--- program side_paint (robot ABB IRB 5500-27) ---
  Smooth(1)
  Set speed (1000.0 mm/s)
  Set Ref.: FrameSidePaint
  Set Tool: Paint gun
  Show Paint gun
  MoveJ 1 to (-1297.14, 952.77, 801.05) mm, rotated rx -98.58 ry 36.73 rz 174.5 deg; joints [-13.501, 53.284, -35.7, -53.192, 43.737, -41.413, -170]
  MoveL 2 to (-1297.14, 952.77, 801.05) mm, rotated rx -98.58 ry 36.73 rz 174.5 deg; joints [-13.501, 53.284, -35.7, -53.192, 43.737, -41.413, -170]
  MoveL 3 to (-1297.75, 853.49, 789.09) mm, rotated rx -98.58 ry 36.73 rz 174.5 deg; joints [-15.474, 56.036, -39.978, -51.479, 40.206, -40.518, -170]
  MoveL 4 to (-1297.75, 853.49, 789.09) mm, rotated rx -98.58 ry 36.73 rz 174.5 deg; joints [-15.474, 56.036, -39.978, -51.479, 40.206, -40.518, -170]
  Set speed (50.0 mm/s)
  MoveL 5 to (-1297.75, 853.39, 796.9) mm, rotated rx -98.58 ry 36.73 rz 174.5 deg; joints [-15.482, 55.905, -40.062, -50.968, 39.758, -40.731, -170]
  Set speed (1000.0 mm/s)
  MoveL 6 to (-1297.75, 853.39, 796.9) mm, rotated rx -98.58 ry 36.73 rz 174.5 deg; joints [-15.482, 55.905, -40.062, -50.968, 39.758, -40.731, -170]
  MoveL 7 to (-1297.14, 952.67, 808.86) mm, rotated rx -98.58 ry 36.73 rz 174.5 deg; joints [-13.509, 53.15, -35.783, -52.711, 43.305, -41.606, -170]
  Set speed (1000.0 mm/s)
  MoveL 8 to (-1377.47, 943.1, 874.94) mm, rotated rx -98.65 ry 38.29 rz 174.46 deg; joints [-14.496, 49.055, -31.026, -57.58, 47.073, -38.423, -170]
  MoveL 9 to (-1377.75, 843.8, 863.14) mm, rotated rx -98.65 ry 38.29 rz 174.46 deg; joints [-16.488, 51.747, -35.093, -56.497, 44.013, -37.161, -170]
  MoveL 10 to (-1377.75, 843.8, 863.14) mm, rotated rx -98.65 ry 38.29 rz 174.46 deg; joints [-16.488, 51.747, -35.093, -56.497, 44.013, -37.161, -170]
  Set speed (50.0 mm/s)
  MoveL 11 to (-1377.75, 845.82, 854.57) mm, rotated rx -98.73 ry 37.85 rz 174.4 deg; joints [-16.458, 51.746, -34.877, -56.091, 43.595, -37.432, -170]
  MoveL 12 to (-1377.75, 852.68, 825.37) mm, rotated rx -98.99 ry 36.5 rz 174.23 deg; joints [-16.347, 51.788, -34.184, -54.959, 42.475, -38.231, -170]
  MoveL 13 to (-1377.75, 852.68, 825.37) mm, rotated rx -98.99 ry 36.5 rz 174.23 deg; joints [-16.347, 51.788, -34.184, -54.959, 42.475, -38.231, -170]
  MoveL 14 to (-1377.75, 852.9, 804.32) mm, rotated rx -98.93 ry 36.57 rz 174.27 deg; joints [-16.325, 52.17, -33.954, -56.498, 43.866, -37.653, -170]
  MoveL 15 to (-1377.75, 853.2, 774.32) mm, rotated rx -98.85 ry 36.66 rz 174.33 deg; joints [-16.297, 52.733, -33.656, -58.588, 45.794, -36.9, -170]
  MoveL 16 to (-1377.75, 853.51, 744.32) mm, rotated rx -98.76 ry 36.76 rz 174.38 deg; joints [-16.27, 53.316, -33.393, -60.572, 47.664, -36.222, -170]
  MoveL 17 to (-1377.75, 853.62, 723.27) mm, rotated rx -96.67 ry 38.01 rz 175.72 deg; joints [-16.272, 54.302, -33.281, -66.947, 53.226, -34.784, -170]
  MoveL 18 to (-1377.75, 853.79, 693.27) mm, rotated rx -92.96 ry 22.32 rz 178.98 deg; joints [-17.183, 52.483, -31.27, -47.624, 27.861, -47.672, -170]
  MoveL 19 to (-1377.75, 853.95, 663.27) mm, rotated rx -90.24 ry 20.37 rz -179.71 deg; joints [-17.303, 53.259, -30.78, -52.353, 29.913, -47.74, -170]
  MoveL 20 to (-1377.75, 854, 636.95) mm, rotated rx -90.22 ry 20.39 rz -179.69 deg; joints [-17.278, 53.814, -30.63, -54.436, 31.655, -46.867, -170]
  MoveL 21 to (-1377.75, 854.06, 606.95) mm, rotated rx -90.19 ry 20.4 rz -179.67 deg; joints [-17.254, 54.461, -30.491, -56.636, 33.537, -45.983, -170]
  MoveL 22 to (-1377.75, 854.12, 576.95) mm, rotated rx -90.16 ry 20.41 rz -179.64 deg; joints [-17.232, 55.127, -30.383, -58.679, 35.325, -45.201, -170]
  MoveL 23 to (-1377.75, 854.18, 546.95) mm, rotated rx -90.13 ry 20.43 rz -179.62 deg; joints [-17.213, 55.809, -30.307, -60.585, 37.031, -44.505, -170]
  MoveL 24 to (-1377.75, 854.23, 516.95) mm, rotated rx -90.1 ry 20.44 rz -179.6 deg; joints [-17.195, 56.507, -30.263, -62.373, 38.664, -43.883, -170]
  MoveL 25 to (-1377.75, 854.25, 508.95) mm, rotated rx -90.1 ry 20.44 rz -179.6 deg; joints [-17.19, 56.695, -30.258, -62.801, 39.067, -43.739, -170]
  Set speed (1000.0 mm/s)
  MoveL 26 to (-1377.75, 854.25, 508.95) mm, rotated rx -90.1 ry 20.44 rz -179.6 deg; joints [-17.19, 56.695, -30.258, -62.801, 39.067, -43.739, -170]
  MoveL 27 to (-1378.51, 954.25, 509.11) mm, rotated rx -90.1 ry 20.44 rz -179.6 deg; joints [-15.183, 54.375, -26.133, -63.747, 42.417, -45.012, -170]
  Set speed (1000.0 mm/s)
  MoveL 28 to (-1458.68, 953.67, 187.25) mm, rotated rx -89.99 ry 0.54 rz -179.47 deg; joints [-16.728, 56.853, -21.556, -35.057, 15.198, -66.186, -170]
  MoveL 29 to (-1457.75, 853.67, 187.27) mm, rotated rx -89.99 ry 0.54 rz -179.47 deg; joints [-18.915, 58.968, -25.635, -25.442, 6.373, -70.654, -170]
  MoveL 30 to (-1457.75, 853.67, 187.27) mm, rotated rx -89.99 ry 0.54 rz -179.47 deg; joints [-18.915, 58.968, -25.635, -25.442, 6.373, -70.654, -170]
  Set speed (50.0 mm/s)
  MoveL 31 to (-1457.75, 853.67, 195.27) mm, rotated rx -89.99 ry 0.54 rz -179.47 deg; joints [-18.972, 58.745, -25.612, -22.234, 4.29, -72.531, -170]
  MoveL 32 to (-1457.75, 853.67, 225.27) mm, rotated rx -90 ry 20.52 rz -179.48 deg; joints [-18.06, 61.359, -26.112, -80.802, 56.365, -38.648, -170]
  MoveL 33 to (-1457.75, 853.67, 255.27) mm, rotated rx -90 ry 20.51 rz -179.49 deg; joints [-18.066, 60.5, -25.864, -79.807, 55.247, -38.783, -170]
  MoveL 34 to (-1457.75, 853.67, 285.27) mm, rotated rx -90.01 ry 20.51 rz -179.5 deg; joints [-18.073, 59.656, -25.644, -78.771, 54.095, -38.938, -170]
  MoveL 35 to (-1457.75, 853.67, 315.27) mm, rotated rx -90.01 ry 20.5 rz -179.51 deg; joints [-18.079, 58.826, -25.455, -77.693, 52.908, -39.114, -170]
  MoveL 36 to (-1457.75, 853.67, 345.27) mm, rotated rx -90.02 ry 20.49 rz -179.52 deg; joints [-18.087, 58.011, -25.294, -76.57, 51.684, -39.312, -170]
  MoveL 37 to (-1457.75, 853.67, 375.27) mm, rotated rx -90.02 ry 20.48 rz -179.53 deg; joints [-18.095, 57.21, -25.164, -75.399, 50.423, -39.536, -170]
  MoveL 38 to (-1457.75, 853.66, 405.27) mm, rotated rx -90.03 ry 20.48 rz -179.53 deg; joints [-18.104, 56.424, -25.062, -74.178, 49.125, -39.788, -170]
  MoveL 39 to (-1457.75, 853.66, 435.27) mm, rotated rx -90.03 ry 20.47 rz -179.54 deg; joints [-18.114, 55.652, -24.99, -72.903, 47.786, -40.071, -170]
  MoveL 40 to (-1457.75, 853.66, 465.27) mm, rotated rx -90.04 ry 20.46 rz -179.55 deg; joints [-18.124, 54.896, -24.946, -71.569, 46.405, -40.387, -170]
  MoveL 41 to (-1457.75, 853.66, 495.27) mm, rotated rx -90.04 ry 20.46 rz -179.56 deg; joints [-18.135, 54.155, -24.932, -70.172, 44.981, -40.741, -170]
  MoveL 42 to (-1457.75, 853.66, 526.08) mm, rotated rx -90.05 ry 20.45 rz -179.57 deg; joints [-18.148, 53.41, -24.949, -68.666, 43.469, -41.147, -170]
  MoveL 43 to (-1457.75, 853.62, 556.08) mm, rotated rx -90.07 ry 20.43 rz -179.59 deg; joints [-18.161, 52.696, -24.998, -67.057, 41.898, -41.604, -170]
  MoveL 44 to (-1457.75, 853.58, 586.08) mm, rotated rx -90.1 ry 20.42 rz -179.62 deg; joints [-18.176, 51.999, -25.077, -65.36, 40.27, -42.117, -170]
  MoveL 45 to (-1457.75, 853.52, 628.44) mm, rotated rx -90.14 ry 20.4 rz -179.65 deg; joints [-18.199, 51.042, -25.24, -62.791, 37.864, -42.951, -170]
  MoveL 46 to (-1457.75, 853.41, 658.44) mm, rotated rx -90.2 ry 20.38 rz -179.69 deg; joints [-18.219, 50.379, -25.397, -60.74, 36.008, -43.651, -170]
  MoveL 47 to (-1457.75, 853.3, 688.44) mm, rotated rx -90.25 ry 20.36 rz -179.73 deg; joints [-18.241, 49.734, -25.586, -58.544, 34.065, -44.447, -170]
  MoveL 48 to (-1457.75, 853.15, 730.8) mm, rotated rx -90.34 ry 20.33 rz -179.78 deg; joints [-18.277, 48.852, -25.907, -55.141, 31.145, -45.766, -170]
  MoveL 49 to (-1457.75, 852.89, 760.79) mm, rotated rx -92.62 ry 22.9 rz 179.1 deg; joints [-18.125, 48.27, -26.437, -53.114, 31.255, -44.471, -170]
  MoveL 50 to (-1457.75, 852.62, 790.79) mm, rotated rx -94.76 ry 18.59 rz 178.38 deg; joints [-18.675, 46.691, -27.128, -19.032, 6.195, -62.515, -170]
  MoveL 51 to (-1457.75, 852.24, 833.15) mm, rotated rx -99.29 ry 36.39 rz 174.04 deg; joints [-17.25, 48.344, -28.68, -59.788, 46.031, -35.543, -170]
  MoveL 52 to (-1457.75, 842.15, 874) mm, rotated rx -99.06 ry 37.76 rz 174.19 deg; joints [-17.436, 48.149, -29.605, -60.089, 46.37, -34.987, -170]
  MoveL 53 to (-1457.75, 832.57, 914.98) mm, rotated rx -98.75 ry 39.5 rz 174.39 deg; joints [-17.596, 48.056, -30.593, -61.046, 47.459, -34.165, -170]
  MoveL 54 to (-1457.75, 829.64, 928.8) mm, rotated rx -100.09 ry 40.17 rz 173.53 deg; joints [-17.613, 47.828, -31.021, -59.139, 46.443, -34.036, -170]
  Set speed (1000.0 mm/s)
  MoveL 55 to (-1457.75, 829.64, 928.8) mm, rotated rx -100.09 ry 40.17 rz 173.53 deg; joints [-17.613, 47.828, -31.021, -59.139, 46.443, -34.036, -170]
  MoveL 56 to (-1457.88, 928.74, 942.19) mm, rotated rx -100.09 ry 40.17 rz 173.53 deg; joints [-15.61, 45.122, -27.108, -59.778, 49.118, -35.52, -170]
  Set speed (1000.0 mm/s)
  MoveL 57 to (-1538.66, 913.21, 1014.54) mm, rotated rx -105.61 ry 41.62 rz 170.03 deg; joints [-16.814, 40.69, -24.051, -54.13, 45.376, -33.626, -170]
  MoveL 58 to (-1537.75, 815.25, 994.43) mm, rotated rx -105.61 ry 41.62 rz 170.03 deg; joints [-18.805, 43.502, -27.729, -53.938, 43.177, -32.043, -170]
  MoveL 59 to (-1537.75, 815.25, 994.43) mm, rotated rx -105.61 ry 41.62 rz 170.03 deg; joints [-18.805, 43.502, -27.729, -53.938, 43.177, -32.043, -170]
  Set speed (50.0 mm/s)
  MoveL 60 to (-1537.75, 817.42, 984.35) mm, rotated rx -105.7 ry 41.25 rz 169.97 deg; joints [-18.767, 43.525, -27.488, -53.735, 42.978, -32.204, -170]
  MoveL 61 to (-1537.75, 823.74, 955.02) mm, rotated rx -106.39 ry 38.88 rz 169.55 deg; joints [-18.708, 43.372, -26.899, -49.424, 39.023, -34.352, -170]
  MoveL 62 to (-1537.75, 830.36, 927.04) mm, rotated rx -102.94 ry 38.8 rz 171.73 deg; joints [-18.566, 44.073, -25.879, -57.39, 44.7, -32.92, -170]
  MoveL 63 to (-1537.75, 837.26, 897.85) mm, rotated rx -99.3 ry 38.2 rz 174.04 deg; joints [-18.489, 44.817, -24.916, -64.229, 49.447, -32.46, -170]
  MoveL 64 to (-1537.75, 844.38, 869.99) mm, rotated rx -99.44 ry 37.24 rz 173.95 deg; joints [-18.359, 44.951, -24.277, -64.056, 49.208, -32.848, -170]
  MoveL 65 to (-1537.75, 851.81, 840.93) mm, rotated rx -108.52 ry 36.78 rz 168.22 deg; joints [-18.104, 43.97, -24.492, -49.321, 40.009, -34.298, -170]
  MoveL 66 to (-1537.75, 852.15, 797.55) mm, rotated rx -101.05 ry 38.75 rz 172.92 deg; joints [-18.073, 46.114, -23.379, -67.854, 54.496, -30.798, -170]
  MoveL 67 to (-1537.75, 852.4, 767.56) mm, rotated rx -94.65 ry 21.55 rz 178.41 deg; joints [-19.181, 44.634, -21.632, -51.982, 29.331, -43.354, -170]
  MoveL 68 to (-1537.75, 852.64, 737.56) mm, rotated rx -90.09 ry 20.34 rz -179.69 deg; joints [-19.27, 45.923, -20.99, -62.422, 36.243, -42.294, -170]
  MoveL 69 to (-1537.75, 852.77, 694.18) mm, rotated rx -90.06 ry 20.37 rz -179.66 deg; joints [-19.242, 46.844, -20.673, -65.334, 38.948, -41.323, -170]
  MoveL 70 to (-1537.75, 852.86, 664.18) mm, rotated rx -90.04 ry 20.38 rz -179.63 deg; joints [-19.226, 47.501, -20.49, -67.203, 40.732, -40.746, -170]
  MoveL 71 to (-1537.75, 852.95, 634.18) mm, rotated rx -90.02 ry 20.4 rz -179.6 deg; joints [-19.211, 48.176, -20.337, -68.97, 42.453, -40.235, -170]
  MoveL 72 to (-1537.75, 852.98, 590.81) mm, rotated rx -90 ry 20.42 rz -179.58 deg; joints [-19.193, 49.178, -20.172, -71.312, 44.799, -39.612, -170]
  MoveL 73 to (-1537.75, 853.01, 560.81) mm, rotated rx -89.99 ry 20.44 rz -179.56 deg; joints [-19.181, 49.891, -20.094, -72.839, 46.362, -39.24, -170]
  MoveL 74 to (-1537.75, 853.03, 530.81) mm, rotated rx -89.98 ry 20.45 rz -179.55 deg; joints [-19.171, 50.619, -20.044, -74.297, 47.879, -38.91, -170]
  MoveL 75 to (-1537.75, 853.02, 496.12) mm, rotated rx -89.98 ry 20.46 rz -179.54 deg; joints [-19.16, 51.478, -20.025, -75.864, 49.547, -38.588, -170]
  MoveL 76 to (-1537.75, 853.02, 466.12) mm, rotated rx -89.98 ry 20.47 rz -179.53 deg; joints [-19.151, 52.238, -20.038, -77.16, 50.948, -38.345, -170]
  MoveL 77 to (-1537.75, 853.01, 436.12) mm, rotated rx -89.97 ry 20.47 rz -179.52 deg; joints [-19.143, 53.012, -20.08, -78.405, 52.311, -38.132, -170]
  MoveL 78 to (-1537.75, 853, 406.12) mm, rotated rx -89.97 ry 20.48 rz -179.51 deg; joints [-19.136, 53.8, -20.15, -79.602, 53.639, -37.945, -170]
  MoveL 79 to (-1537.75, 852.99, 376.12) mm, rotated rx -89.97 ry 20.49 rz -179.51 deg; joints [-19.129, 54.603, -20.249, -80.755, 54.932, -37.784, -170]
  MoveL 80 to (-1537.75, 852.98, 346.12) mm, rotated rx -89.97 ry 20.49 rz -179.5 deg; joints [-19.123, 55.42, -20.375, -81.866, 56.191, -37.645, -170]
  MoveL 81 to (-1537.75, 852.97, 316.12) mm, rotated rx -89.97 ry 20.5 rz -179.49 deg; joints [-19.117, 56.251, -20.529, -82.938, 57.418, -37.526, -170]
  MoveL 82 to (-1537.75, 852.96, 286.12) mm, rotated rx -89.97 ry 0.51 rz -179.49 deg; joints [-19.911, 53.732, -20.278, -31.164, 8.952, -66.908, -170]
  MoveL 83 to (-1537.75, 852.95, 256.12) mm, rotated rx -89.97 ry 0.52 rz -179.49 deg; joints [-19.811, 54.549, -20.328, -37.182, 13.072, -63.574, -170]
  MoveL 84 to (-1537.75, 852.94, 226.12) mm, rotated rx -89.97 ry 0.52 rz -179.48 deg; joints [-19.743, 55.38, -20.423, -41.507, 16.152, -61.281, -170]
  MoveL 85 to (-1537.75, 852.94, 196.12) mm, rotated rx -89.97 ry 0.53 rz -179.47 deg; joints [-19.691, 56.224, -20.555, -44.993, 18.721, -59.506, -170]
  MoveL 86 to (-1537.75, 852.93, 188.12) mm, rotated rx -89.97 ry 0.53 rz -179.47 deg; joints [-19.679, 56.452, -20.597, -45.807, 19.336, -59.104, -170]
  Set speed (1000.0 mm/s)
  MoveL 87 to (-1537.75, 852.93, 188.12) mm, rotated rx -89.97 ry 0.53 rz -179.47 deg; joints [-19.679, 56.452, -20.597, -45.807, 19.336, -59.104, -170]
  MoveL 88 to (-1538.66, 952.93, 188.06) mm, rotated rx -89.97 ry 0.53 rz -179.47 deg; joints [-17.579, 54.397, -16.722, -48.142, 23.689, -59.07, -170]
  Set speed (1000.0 mm/s)
  MoveL 89 to (-1618.68, 952.19, 188.9) mm, rotated rx -89.96 ry 0.54 rz -179.47 deg; joints [-18.571, 52.085, -12.202, -57.393, 29.915, -54.439, -170]
  MoveL 90 to (-1617.75, 852.2, 188.97) mm, rotated rx -89.96 ry 0.54 rz -179.47 deg; joints [-20.682, 54.098, -15.965, -56.732, 26.603, -53.482, -170]
  MoveL 91 to (-1617.75, 852.2, 188.97) mm, rotated rx -89.96 ry 0.54 rz -179.47 deg; joints [-20.682, 54.098, -15.965, -56.732, 26.603, -53.482, -170]
  Set speed (50.0 mm/s)
  MoveL 92 to (-1617.75, 852.2, 196.97) mm, rotated rx -89.96 ry 0.54 rz -179.47 deg; joints [-20.69, 53.866, -15.922, -56.157, 26.118, -53.721, -170]
  MoveL 93 to (-1617.75, 852.22, 226.97) mm, rotated rx -89.97 ry 0.52 rz -179.48 deg; joints [-20.719, 53.003, -15.784, -53.748, 24.141, -54.766, -170]
  MoveL 94 to (-1617.75, 852.24, 256.97) mm, rotated rx -89.97 ry 0.52 rz -179.49 deg; joints [-20.754, 52.154, -15.675, -51.107, 22.023, -55.958, -170]
  MoveL 95 to (-1617.75, 852.26, 286.97) mm, rotated rx -89.97 ry 0.51 rz -179.49 deg; joints [-20.796, 51.317, -15.598, -48.095, 19.679, -57.38, -170]
  MoveL 96 to (-1617.75, 852.27, 316.97) mm, rotated rx -89.97 ry 0.5 rz -179.5 deg; joints [-20.847, 50.495, -15.554, -44.557, 17.016, -59.128, -170]
  MoveL 97 to (-1617.75, 852.29, 346.97) mm, rotated rx -89.97 ry 0.5 rz -179.51 deg; joints [-20.914, 49.687, -15.548, -40.195, 13.853, -61.388, -170]
  MoveL 98 to (-1617.75, 852.31, 376.97) mm, rotated rx -89.98 ry 0.49 rz -179.51 deg; joints [-21.012, 48.892, -15.587, -34.212, 9.696, -64.645, -170]
  MoveL 99 to (-1617.75, 852.33, 406.97) mm, rotated rx -89.98 ry 20.48 rz -179.51 deg; joints [-20.237, 51.333, -15.572, -84.454, 57.702, -36.409, -170]
  MoveL 100 to (-1617.75, 852.35, 436.97) mm, rotated rx -89.98 ry 20.47 rz -179.52 deg; joints [-20.242, 50.524, -15.503, -83.301, 56.367, -36.513, -170]
  MoveL 101 to (-1617.75, 852.37, 466.97) mm, rotated rx -89.98 ry 20.47 rz -179.53 deg; joints [-20.248, 49.73, -15.463, -82.109, 55.001, -36.64, -170]
  MoveL 102 to (-1617.75, 852.39, 496.97) mm, rotated rx -89.98 ry 20.46 rz -179.54 deg; joints [-20.255, 48.951, -15.449, -80.875, 53.602, -36.792, -170]
  MoveL 103 to (-1617.75, 852.41, 535.54) mm, rotated rx -89.98 ry 20.45 rz -179.55 deg; joints [-20.264, 47.97, -15.472, -79.22, 51.753, -37.028, -170]
  MoveL 104 to (-1617.75, 852.4, 565.54) mm, rotated rx -90.01 ry 20.44 rz -179.57 deg; joints [-20.271, 47.22, -15.523, -77.823, 50.231, -37.252, -170]
  MoveL 105 to (-1617.75, 852.39, 595.54) mm, rotated rx -90.03 ry 20.42 rz -179.59 deg; joints [-20.279, 46.485, -15.603, -76.37, 48.67, -37.512, -170]
  MoveL 106 to (-1617.75, 852.38, 639.93) mm, rotated rx -90.06 ry 20.41 rz -179.62 deg; joints [-20.293, 45.427, -15.772, -74.103, 46.282, -37.971, -170]
  MoveL 107 to (-1617.75, 852.31, 669.93) mm, rotated rx -90.12 ry 20.39 rz -179.65 deg; joints [-20.304, 44.727, -15.926, -72.412, 44.555, -38.344, -170]
  MoveL 108 to (-1617.75, 852.24, 699.93) mm, rotated rx -90.17 ry 20.37 rz -179.69 deg; joints [-20.316, 44.043, -16.108, -70.636, 42.774, -38.773, -170]
  MoveL 109 to (-1617.75, 852.13, 744.32) mm, rotated rx -90.25 ry 20.34 rz -179.74 deg; joints [-20.337, 43.062, -16.432, -67.828, 40.03, -39.528, -170]
  MoveL 110 to (-1617.75, 851.91, 774.32) mm, rotated rx -92.66 ry 22.74 rz 179.08 deg; joints [-20.17, 42.355, -16.931, -65.107, 39.405, -38.293, -170]
  MoveL 111 to (-1617.75, 851.69, 804.32) mm, rotated rx -94.93 ry 18.43 rz 178.32 deg; joints [-20.429, 40.696, -17.575, -45.711, 22.412, -46.525, -170]
  MoveL 112 to (-1617.75, 851.37, 848.7) mm, rotated rx -99.89 ry 36.19 rz 173.66 deg; joints [-19.251, 42.062, -18.981, -67.544, 51.608, -31.157, -170]
  MoveL 113 to (-1617.75, 843.67, 877.7) mm, rotated rx -99.76 ry 37.11 rz 173.74 deg; joints [-19.4, 41.875, -19.608, -67.602, 51.704, -30.786, -170]
  MoveL 114 to (-1617.75, 834.4, 912.57) mm, rotated rx -99.62 ry 38.3 rz 173.84 deg; joints [-19.573, 41.685, -20.402, -67.708, 51.904, -30.316, -170]
  MoveL 115 to (-1617.75, 827.27, 941.71) mm, rotated rx -102.97 ry 39.03 rz 171.7 deg; joints [-19.648, 40.983, -21.342, -61.801, 47.743, -30.345, -170]
  MoveL 116 to (-1617.75, 818.68, 976.75) mm, rotated rx -106.97 ry 39.25 rz 169.19 deg; joints [-19.823, 40.144, -22.589, -53.1, 41.333, -31.482, -170]
  MoveL 117 to (-1617.75, 812.22, 1006.05) mm, rotated rx -106.44 ry 40.96 rz 169.51 deg; joints [-19.915, 40.172, -23.197, -55.546, 43.623, -30.225, -170]
  MoveL 118 to (-1617.75, 807.51, 1027.38) mm, rotated rx -106.08 ry 42.33 rz 169.72 deg; joints [-19.975, 40.225, -23.674, -57.365, 45.437, -29.299, -170]
  Set speed (1000.0 mm/s)
  MoveL 119 to (-1617.75, 807.51, 1027.38) mm, rotated rx -106.08 ry 42.33 rz 169.72 deg; joints [-19.975, 40.225, -23.674, -57.365, 45.437, -29.299, -170]
  MoveL 120 to (-1618.95, 905.38, 1047.86) mm, rotated rx -106.08 ry 42.33 rz 169.72 deg; joints [-17.969, 37.4, -20.103, -57.146, 47.301, -31.08, -170]
  Set speed (1000.0 mm/s)
  MoveL 121 to (-1698.82, 903.07, 1054.33) mm, rotated rx -106.93 ry 41.66 rz 169.19 deg; joints [-19.102, 34.266, -15.907, -58.357, 47.41, -29.419, -170]
  MoveL 122 to (-1697.75, 805.47, 1032.58) mm, rotated rx -106.93 ry 41.66 rz 169.19 deg; joints [-21.13, 37.101, -19.331, -59.044, 45.923, -27.455, -170]
  MoveL 123 to (-1697.75, 805.47, 1032.58) mm, rotated rx -106.93 ry 41.66 rz 169.19 deg; joints [-21.13, 37.101, -19.331, -59.044, 45.923, -27.455, -170]
  Set speed (50.0 mm/s)
  MoveL 124 to (-1697.75, 810.24, 1012.22) mm, rotated rx -106.94 ry 41.63 rz 169.19 deg; joints [-21.016, 37.286, -18.807, -60.335, 47.246, -27.094, -170]
  MoveL 125 to (-1697.75, 817.08, 983.01) mm, rotated rx -107.81 ry 38.8 rz 168.66 deg; joints [-20.955, 37.062, -18.305, -55.172, 42.194, -29.411, -170]
  MoveL 126 to (-1697.75, 825.95, 948.64) mm, rotated rx -103.6 ry 38.71 rz 171.31 deg; joints [-20.77, 37.953, -17.013, -64.34, 49.163, -28.359, -170]
  MoveL 127 to (-1697.75, 833.44, 919.6) mm, rotated rx -99.99 ry 38.1 rz 173.6 deg; joints [-20.691, 38.726, -16.038, -70.745, 53.9, -28.428, -170]
  MoveL 128 to (-1697.75, 842.92, 885.39) mm, rotated rx -100.1 ry 36.99 rz 173.53 deg; joints [-20.509, 38.936, -15.26, -70.769, 53.836, -28.878, -170]
  MoveL 129 to (-1697.75, 850.93, 856.48) mm, rotated rx -100.2 ry 36.09 rz 173.46 deg; joints [-20.351, 39.14, -14.634, -70.808, 53.837, -29.243, -170]
  MoveL 130 to (-1697.75, 851.03, 841.08) mm, rotated rx -97.37 ry 16.83 rz 177.49 deg; joints [-21.807, 36.737, -14.224, -31.988, 11.526, -51.964, -170]
  MoveL 131 to (-1697.75, 851.23, 811.08) mm, rotated rx -95.02 ry 18.35 rz 178.29 deg; joints [-21.516, 37.902, -13.293, -52.995, 26.817, -42.288, -170]
  MoveL 132 to (-1697.75, 851.43, 781.08) mm, rotated rx -92.69 ry 22.66 rz 179.07 deg; joints [-21.307, 39.604, -12.646, -69.982, 42.691, -35.881, -170]
  MoveL 133 to (-1697.75, 851.63, 751.08) mm, rotated rx -90.21 ry 20.35 rz -179.73 deg; joints [-21.485, 40.373, -12.157, -72.974, 43.653, -37.152, -170]
  MoveL 134 to (-1697.75, 851.65, 735.67) mm, rotated rx -90.18 ry 20.36 rz -179.71 deg; joints [-21.479, 40.719, -12.038, -73.897, 44.596, -36.946, -170]
  MoveL 135 to (-1697.75, 851.7, 705.67) mm, rotated rx -90.13 ry 20.37 rz -179.67 deg; joints [-21.469, 41.405, -11.828, -75.631, 46.392, -36.59, -170]
  MoveL 136 to (-1697.75, 851.76, 675.67) mm, rotated rx -90.08 ry 20.39 rz -179.64 deg; joints [-21.46, 42.108, -11.646, -77.288, 48.141, -36.285, -170]
  MoveL 137 to (-1697.75, 851.81, 645.67) mm, rotated rx -90.03 ry 20.41 rz -179.6 deg; joints [-21.452, 42.828, -11.492, -78.876, 49.844, -36.028, -170]
  MoveL 138 to (-1697.75, 851.8, 630.27) mm, rotated rx -90.02 ry 20.41 rz -179.59 deg; joints [-21.448, 43.201, -11.426, -79.634, 50.676, -35.912, -170]
  MoveL 139 to (-1697.75, 851.8, 600.27) mm, rotated rx -90 ry 20.43 rz -179.57 deg; joints [-21.442, 43.94, -11.318, -81.07, 52.266, -35.714, -170]
  MoveL 140 to (-1697.75, 851.79, 570.27) mm, rotated rx -89.98 ry 20.44 rz -179.55 deg; joints [-21.436, 44.694, -11.238, -82.453, 53.821, -35.549, -170]
  MoveL 141 to (-1697.75, 851.78, 540.27) mm, rotated rx -89.96 ry 20.45 rz -179.53 deg; joints [-21.431, 45.464, -11.184, -83.789, 55.341, -35.415, -170]
  MoveL 142 to (-1697.75, 851.74, 497.81) mm, rotated rx -89.95 ry 20.46 rz -179.52 deg; joints [-21.424, 46.572, -11.158, -85.539, 57.381, -35.274, -170]
  MoveL 143 to (-1697.75, 851.72, 467.81) mm, rotated rx -89.96 ry 0.47 rz -179.53 deg; joints [-22.229, 44.199, -11.448, -34.327, 8.364, -63.992, -170]
  MoveL 144 to (-1697.75, 851.69, 437.81) mm, rotated rx -89.96 ry 0.48 rz -179.53 deg; joints [-22.114, 44.971, -11.312, -41.283, 13.178, -60.192, -170]
  MoveL 145 to (-1697.75, 851.66, 407.81) mm, rotated rx -89.96 ry 0.48 rz -179.52 deg; joints [-22.04, 45.758, -11.23, -46.061, 16.652, -57.729, -170]
  MoveL 146 to (-1697.75, 851.63, 377.81) mm, rotated rx -89.96 ry 0.49 rz -179.51 deg; joints [-21.985, 46.558, -11.187, -49.857, 19.528, -55.875, -170]
  MoveL 147 to (-1697.75, 851.6, 347.81) mm, rotated rx -89.95 ry 0.5 rz -179.51 deg; joints [-21.941, 47.374, -11.179, -53.056, 22.044, -54.391, -170]
  MoveL 148 to (-1697.75, 851.58, 317.81) mm, rotated rx -89.95 ry 0.5 rz -179.5 deg; joints [-21.904, 48.203, -11.203, -55.845, 24.311, -53.164, -170]
  MoveL 149 to (-1697.75, 851.55, 287.81) mm, rotated rx -89.95 ry 0.51 rz -179.49 deg; joints [-21.874, 49.046, -11.258, -58.327, 26.391, -52.127, -170]
  MoveL 150 to (-1697.75, 851.52, 257.81) mm, rotated rx -89.95 ry 0.52 rz -179.49 deg; joints [-21.847, 49.902, -11.343, -60.569, 28.324, -51.239, -170]
  MoveL 151 to (-1697.75, 851.49, 227.81) mm, rotated rx -89.95 ry 0.52 rz -179.48 deg; joints [-21.825, 50.772, -11.458, -62.618, 30.136, -50.47, -170]
  MoveL 152 to (-1697.75, 851.46, 197.81) mm, rotated rx -89.95 ry 0.53 rz -179.47 deg; joints [-21.804, 51.654, -11.602, -64.505, 31.847, -49.8, -170]
  MoveL 153 to (-1697.75, 851.46, 189.81) mm, rotated rx -89.95 ry 0.53 rz -179.47 deg; joints [-21.799, 51.892, -11.646, -64.974, 32.281, -49.642, -170]
  Set speed (1000.0 mm/s)
  MoveL 154 to (-1697.75, 851.46, 189.81) mm, rotated rx -89.95 ry 0.53 rz -179.47 deg; joints [-21.799, 51.892, -11.646, -64.974, 32.281, -49.642, -170]
  MoveL 155 to (-1698.67, 951.45, 189.73) mm, rotated rx -89.95 ry 0.53 rz -179.47 deg; joints [-19.662, 49.906, -7.955, -64.826, 35.07, -51.053, -170]
  Set speed (1000.0 mm/s)
  MoveL 156 to (-1778.68, 950.71, 190.56) mm, rotated rx -89.94 ry 0.54 rz -179.46 deg; joints [-20.852, 47.841, -3.934, -71.319, 39.653, -48.345, -170]
  MoveL 157 to (-1777.75, 850.72, 190.66) mm, rotated rx -89.94 ry 0.54 rz -179.46 deg; joints [-23.016, 49.811, -7.581, -71.951, 37.192, -46.68, -170]
  MoveL 158 to (-1777.75, 850.72, 190.66) mm, rotated rx -89.94 ry 0.54 rz -179.46 deg; joints [-23.016, 49.811, -7.581, -71.951, 37.192, -46.68, -170]
  Set speed (50.0 mm/s)
  MoveL 159 to (-1777.75, 850.73, 198.66) mm, rotated rx -89.94 ry 0.54 rz -179.46 deg; joints [-23.02, 49.568, -7.536, -71.545, 36.785, -46.785, -170]
  MoveL 160 to (-1777.75, 850.76, 228.66) mm, rotated rx -89.94 ry 0.52 rz -179.48 deg; joints [-23.033, 48.664, -7.392, -69.892, 35.171, -47.256, -170]
  MoveL 161 to (-1777.75, 850.8, 258.66) mm, rotated rx -89.94 ry 0.52 rz -179.48 deg; joints [-23.049, 47.773, -7.274, -68.162, 33.506, -47.774, -170]
  MoveL 162 to (-1777.75, 850.84, 288.66) mm, rotated rx -89.94 ry 0.51 rz -179.49 deg; joints [-23.067, 46.895, -7.184, -66.305, 31.758, -48.368, -170]
  MoveL 163 to (-1777.75, 850.88, 318.66) mm, rotated rx -89.94 ry 0.5 rz -179.5 deg; joints [-23.088, 46.03, -7.122, -64.299, 29.916, -49.054, -170]
  MoveL 164 to (-1777.75, 850.91, 348.66) mm, rotated rx -89.94 ry 0.5 rz -179.5 deg; joints [-23.112, 45.179, -7.09, -62.115, 27.963, -49.85, -170]
  MoveL 165 to (-1777.75, 850.95, 378.66) mm, rotated rx -89.93 ry 0.49 rz -179.51 deg; joints [-23.139, 44.341, -7.087, -59.714, 25.877, -50.78, -170]
  MoveL 166 to (-1777.75, 850.99, 408.66) mm, rotated rx -89.93 ry 0.48 rz -179.52 deg; joints [-23.172, 43.518, -7.115, -57.04, 23.624, -51.882, -170]
  MoveL 167 to (-1777.75, 851.03, 438.66) mm, rotated rx -89.93 ry 0.48 rz -179.52 deg; joints [-23.211, 42.71, -7.175, -54.006, 21.153, -53.208, -170]
  MoveL 168 to (-1777.75, 851.06, 468.66) mm, rotated rx -89.93 ry 0.47 rz -179.53 deg; joints [-23.26, 41.916, -7.268, -50.469, 18.377, -54.848, -170]
  MoveL 169 to (-1777.75, 851.1, 498.66) mm, rotated rx -89.93 ry 0.46 rz -179.54 deg; joints [-23.324, 41.137, -7.4, -46.155, 15.131, -56.971, -170]
  MoveL 170 to (-1777.75, 851.14, 528.66) mm, rotated rx -89.93 ry 0.46 rz -179.54 deg; joints [-23.415, 40.374, -7.577, -40.383, 10.993, -59.993, -170]
  MoveL 171 to (-1777.75, 851.16, 545) mm, rotated rx -89.93 ry 0.45 rz -179.55 deg; joints [-23.493, 39.964, -7.704, -35.827, 7.867, -62.501, -170]
  MoveL 172 to (-1777.75, 851.18, 575) mm, rotated rx -89.95 ry 20.44 rz -179.54 deg; joints [-22.678, 42.282, -7.198, -86.773, 57.141, -34.043, -170]
  MoveL 173 to (-1777.75, 851.2, 605) mm, rotated rx -89.97 ry 20.43 rz -179.56 deg; joints [-22.682, 41.507, -7.28, -85.441, 55.583, -34.123, -170]
  MoveL 174 to (-1777.75, 851.22, 635) mm, rotated rx -89.98 ry 20.42 rz -179.58 deg; joints [-22.686, 40.748, -7.389, -84.064, 53.994, -34.232, -170]
  MoveL 175 to (-1777.75, 851.24, 651.42) mm, rotated rx -90 ry 20.41 rz -179.59 deg; joints [-22.689, 40.339, -7.46, -83.291, 53.11, -34.305, -170]
  MoveL 176 to (-1777.75, 851.2, 681.42) mm, rotated rx -90.04 ry 20.39 rz -179.62 deg; joints [-22.694, 39.599, -7.615, -81.78, 51.416, -34.463, -170]
  MoveL 177 to (-1777.75, 851.17, 711.42) mm, rotated rx -90.09 ry 20.38 rz -179.66 deg; joints [-22.7, 38.876, -7.797, -80.211, 49.684, -34.661, -170]
  MoveL 178 to (-1777.75, 851.14, 741.42) mm, rotated rx -90.14 ry 20.36 rz -179.69 deg; joints [-22.707, 38.17, -8.007, -78.579, 47.912, -34.902, -170]
  MoveL 179 to (-1777.75, 851.12, 757.84) mm, rotated rx -90.17 ry 20.35 rz -179.71 deg; joints [-22.711, 37.791, -8.134, -77.656, 46.923, -35.055, -170]
  MoveL 180 to (-1777.75, 850.94, 787.84) mm, rotated rx -92.71 ry 22.57 rz 179.07 deg; joints [-22.524, 36.96, -8.616, -74.415, 45.623, -33.725, -170]
  MoveL 181 to (-1777.75, 850.76, 817.84) mm, rotated rx -95.12 ry 18.28 rz 178.25 deg; joints [-22.695, 35.212, -9.271, -59.087, 30.456, -38.79, -170]
  MoveL 182 to (-1777.75, 850.58, 847.84) mm, rotated rx -97.53 ry 16.77 rz 177.43 deg; joints [-22.888, 34.008, -10.178, -42.638, 17.67, -45.374, -170]
  MoveL 183 to (-1777.75, 850.49, 864.26) mm, rotated rx -98.85 ry 16.26 rz 176.98 deg; joints [-23.158, 33.436, -10.805, -26.149, 6.515, -53.721, -170]
  MoveL 184 to (-1777.75, 850.49, 864.26) mm, rotated rx -98.85 ry 16.26 rz 176.98 deg; joints [-23.158, 33.436, -10.805, -26.149, 6.515, -53.721, -170]
  MoveL 185 to (-1777.75, 842.16, 893.08) mm, rotated rx -98.73 ry 17.14 rz 177.03 deg; joints [-23.318, 33.226, -11.395, -27.246, 7.128, -52.616, -170]
  MoveL 186 to (-1777.75, 832.44, 926.74) mm, rotated rx -98.59 ry 18.2 rz 177.07 deg; joints [-23.496, 33.009, -12.109, -28.785, 8.045, -51.161, -170]
  MoveL 187 to (-1777.75, 824.59, 955.7) mm, rotated rx -104.22 ry 38.44 rz 170.91 deg; joints [-21.962, 35.048, -12.977, -66.68, 50.356, -26.419, -170]
  MoveL 188 to (-1777.75, 815.43, 989.51) mm, rotated rx -108.66 ry 38.4 rz 168.13 deg; joints [-22.157, 34.109, -14.325, -57.054, 42.833, -27.374, -170]
  MoveL 189 to (-1777.75, 808.21, 1018.63) mm, rotated rx -108.13 ry 39.94 rz 168.45 deg; joints [-22.279, 34.098, -14.906, -59.096, 44.748, -26.34, -170]
  MoveL 190 to (-1777.75, 803.35, 1038.23) mm, rotated rx -107.79 ry 41.05 rz 168.66 deg; joints [-22.356, 34.113, -15.319, -60.499, 46.145, -25.633, -170]
  Set speed (1000.0 mm/s)
  MoveL 191 to (-1777.75, 803.35, 1038.23) mm, rotated rx -107.79 ry 41.05 rz 168.66 deg; joints [-22.356, 34.113, -15.319, -60.499, 46.145, -25.633, -170]
  MoveL 192 to (-1778.69, 900.66, 1061.27) mm, rotated rx -107.79 ry 41.05 rz 168.66 deg; joints [-20.309, 31.245, -12.013, -59.367, 47.266, -27.762, -170]
  Set speed (1000.0 mm/s)
  MoveL 193 to (-1858.63, 898.13, 1068.59) mm, rotated rx -108.65 ry 40.64 rz 168.13 deg; joints [-21.589, 28.342, -8.368, -60.561, 47.245, -25.952, -170]
  MoveL 194 to (-1857.75, 801.12, 1044.32) mm, rotated rx -108.65 ry 40.64 rz 168.13 deg; joints [-23.653, 31.26, -11.582, -62.113, 46.481, -23.674, -170]
  MoveL 195 to (-1857.75, 801.12, 1044.32) mm, rotated rx -108.65 ry 40.64 rz 168.13 deg; joints [-23.653, 31.26, -11.582, -62.113, 46.481, -23.674, -170]
  Set speed (50.0 mm/s)
  MoveL 196 to (-1857.75, 806.11, 1025.28) mm, rotated rx -108.66 ry 40.57 rz 168.12 deg; joints [-23.535, 31.427, -11.075, -63.227, 47.668, -23.415, -170]
  MoveL 197 to (-1857.75, 813.7, 996.25) mm, rotated rx -109.52 ry 38.06 rz 167.6 deg; joints [-23.436, 31.264, -10.612, -58.78, 43.263, -25.344, -170]
  MoveL 198 to (-1857.75, 823.2, 962.87) mm, rotated rx -104.85 ry 38.2 rz 170.52 deg; joints [-23.229, 32.247, -9.197, -68.868, 51.345, -24.494, -170]
  MoveL 199 to (-1857.75, 831.4, 934.01) mm, rotated rx -98.92 ry 18.07 rz 176.96 deg; joints [-24.654, 30.306, -8.348, -39.73, 14.092, -44.065, -170]
  MoveL 200 to (-1857.75, 841.4, 900.77) mm, rotated rx -99.04 ry 17.04 rz 176.92 deg; joints [-24.447, 30.527, -7.617, -39.143, 13.792, -44.981, -170]
  MoveL 201 to (-1857.75, 850.05, 872.04) mm, rotated rx -99.14 ry 16.18 rz 176.89 deg; joints [-24.264, 30.74, -7.006, -38.748, 13.634, -45.699, -170]
  MoveL 202 to (-1857.75, 850.14, 854.6) mm, rotated rx -97.7 ry 16.71 rz 177.38 deg; joints [-24.102, 31.368, -6.379, -50.372, 22.005, -40.584, -170]
  MoveL 203 to (-1857.75, 850.3, 824.6) mm, rotated rx -95.21 ry 18.2 rz 178.22 deg; joints [-23.965, 32.613, -5.479, -64.446, 33.592, -35.738, -170]
  MoveL 204 to (-1857.75, 850.45, 794.6) mm, rotated rx -92.74 ry 22.48 rz 179.06 deg; joints [-23.822, 34.407, -4.811, -78.531, 48.275, -31.741, -170]
  MoveL 205 to (-1857.75, 850.61, 764.6) mm, rotated rx -90.12 ry 20.35 rz -179.69 deg; joints [-24.021, 35.303, -4.335, -82.011, 49.919, -33.152, -170]
  MoveL 206 to (-1857.75, 850.62, 747.17) mm, rotated rx -90.1 ry 20.36 rz -179.67 deg; joints [-24.018, 35.717, -4.199, -82.941, 50.96, -33.051, -170]
  MoveL 207 to (-1857.75, 850.63, 717.17) mm, rotated rx -90.05 ry 20.38 rz -179.64 deg; joints [-24.014, 36.442, -3.988, -84.496, 52.721, -32.91, -170]
  MoveL 208 to (-1857.75, 850.65, 687.17) mm, rotated rx -90.01 ry 20.4 rz -179.61 deg; joints [-24.01, 37.185, -3.805, -85.998, 54.447, -32.807, -170]
  MoveL 209 to (-1857.75, 850.66, 657.17) mm, rotated rx -89.96 ry 20.41 rz -179.57 deg; joints [-24.007, 37.946, -3.648, -87.451, 56.14, -32.739, -170]
  MoveL 210 to (-1857.75, 850.64, 639.73) mm, rotated rx -89.95 ry 20.42 rz -179.56 deg; joints [-24.006, 38.392, -3.572, -88.244, 57.081, -32.71, -170]
  MoveL 211 to (-1857.75, 850.61, 609.73) mm, rotated rx -89.94 ry 0.43 rz -179.57 deg; joints [-24.8, 36.114, -4.241, -39.007, 8.41, -59.988, -170]
  MoveL 212 to (-1857.75, 850.57, 579.73) mm, rotated rx -89.92 ry 0.44 rz -179.56 deg; joints [-24.681, 36.861, -3.963, -46.378, 13.597, -56.064, -170]
  MoveL 213 to (-1857.75, 850.53, 549.73) mm, rotated rx -89.91 ry 0.46 rz -179.55 deg; joints [-24.607, 37.624, -3.747, -51.361, 17.315, -53.603, -170]
  MoveL 214 to (-1857.75, 850.5, 529.51) mm, rotated rx -89.91 ry 0.46 rz -179.54 deg; joints [-24.57, 38.145, -3.629, -54.03, 19.394, -52.357, -170]
  MoveL 215 to (-1857.75, 850.45, 499.51) mm, rotated rx -89.91 ry 0.47 rz -179.53 deg; joints [-24.525, 38.931, -3.484, -57.442, 22.147, -50.848, -170]
  MoveL 216 to (-1857.75, 850.41, 469.51) mm, rotated rx -89.91 ry 0.47 rz -179.53 deg; joints [-24.489, 39.733, -3.373, -60.394, 24.622, -49.627, -170]
  MoveL 217 to (-1857.75, 850.36, 439.51) mm, rotated rx -89.91 ry 0.48 rz -179.52 deg; joints [-24.459, 40.55, -3.294, -63.01, 26.893, -48.616, -170]
  MoveL 218 to (-1857.75, 850.32, 409.51) mm, rotated rx -89.91 ry 0.49 rz -179.52 deg; joints [-24.433, 41.382, -3.245, -65.371, 29.009, -47.765, -170]
  MoveL 219 to (-1857.75, 850.27, 379.51) mm, rotated rx -89.91 ry 0.49 rz -179.51 deg; joints [-24.411, 42.228, -3.226, -67.526, 30.998, -47.043, -170]
  MoveL 220 to (-1857.75, 850.22, 349.51) mm, rotated rx -89.92 ry 0.5 rz -179.5 deg; joints [-24.393, 43.089, -3.235, -69.513, 32.882, -46.425, -170]
  MoveL 221 to (-1857.75, 850.18, 319.51) mm, rotated rx -89.92 ry 0.51 rz -179.5 deg; joints [-24.376, 43.963, -3.273, -71.359, 34.676, -45.894, -170]
  MoveL 222 to (-1857.75, 850.13, 289.51) mm, rotated rx -89.92 ry 0.51 rz -179.49 deg; joints [-24.361, 44.851, -3.339, -73.084, 36.392, -45.436, -170]
  MoveL 223 to (-1857.75, 850.08, 259.51) mm, rotated rx -89.92 ry 0.52 rz -179.48 deg; joints [-24.349, 45.752, -3.433, -74.704, 38.038, -45.042, -170]
  MoveL 224 to (-1857.75, 850.04, 229.51) mm, rotated rx -89.92 ry 0.53 rz -179.48 deg; joints [-24.337, 46.666, -3.554, -76.232, 39.622, -44.703, -170]
  MoveL 225 to (-1857.75, 849.99, 199.51) mm, rotated rx -89.92 ry 0.53 rz -179.47 deg; joints [-24.327, 47.593, -3.702, -77.677, 41.148, -44.412, -170]
  MoveL 226 to (-1857.75, 849.98, 191.51) mm, rotated rx -89.92 ry 0.53 rz -179.47 deg; joints [-24.324, 47.842, -3.747, -78.042, 41.541, -44.346, -170]
  Set speed (1000.0 mm/s)
  MoveL 227 to (-1857.75, 849.98, 191.51) mm, rotated rx -89.92 ry 0.53 rz -179.47 deg; joints [-24.324, 47.842, -3.747, -78.042, 41.541, -44.346, -170]
  MoveL 228 to (-1858.67, 949.97, 191.38) mm, rotated rx -89.92 ry 0.53 rz -179.47 deg; joints [-22.132, 45.878, -0.124, -77.092, 43.775, -46.165, -170]
  Set speed (1000.0 mm/s)
  MoveL 229 to (-1938.68, 949.23, 192.21) mm, rotated rx -89.91 ry 0.54 rz -179.46 deg; joints [-23.513, 44.009, 3.503, -82.478, 47.626, -44.309, -170]
  MoveL 230 to (-1937.75, 849.24, 192.36) mm, rotated rx -89.91 ry 0.54 rz -179.46 deg; joints [-25.73, 45.975, -0.114, -83.65, 45.561, -42.389, -170]
  MoveL 231 to (-1937.75, 849.24, 192.36) mm, rotated rx -89.91 ry 0.54 rz -179.46 deg; joints [-25.73, 45.975, -0.114, -83.65, 45.561, -42.389, -170]
  Set speed (50.0 mm/s)
  MoveL 232 to (-1937.75, 849.25, 200.36) mm, rotated rx -89.91 ry 0.54 rz -179.46 deg; joints [-25.732, 45.72, -0.069, -83.314, 45.176, -42.423, -170]
  MoveL 233 to (-1937.75, 849.31, 230.36) mm, rotated rx -89.91 ry 0.53 rz -179.48 deg; joints [-25.738, 44.769, 0.08, -81.968, 43.674, -42.601, -170]
  MoveL 234 to (-1937.75, 849.36, 260.36) mm, rotated rx -89.91 ry 0.52 rz -179.48 deg; joints [-25.746, 43.831, 0.204, -80.582, 42.138, -42.799, -170]
  MoveL 235 to (-1937.75, 849.42, 290.36) mm, rotated rx -89.9 ry 0.51 rz -179.49 deg; joints [-25.755, 42.906, 0.301, -79.124, 40.552, -43.039, -170]
  MoveL 236 to (-1937.75, 849.47, 320.36) mm, rotated rx -89.9 ry 0.51 rz -179.5 deg; joints [-25.765, 41.993, 0.371, -77.588, 38.911, -43.325, -170]
  MoveL 237 to (-1937.75, 849.53, 350.36) mm, rotated rx -89.9 ry 0.5 rz -179.5 deg; joints [-25.776, 41.094, 0.413, -75.962, 37.209, -43.664, -170]
  MoveL 238 to (-1937.75, 849.59, 380.36) mm, rotated rx -89.9 ry 0.49 rz -179.51 deg; joints [-25.79, 40.209, 0.428, -74.235, 35.44, -44.066, -170]
  MoveL 239 to (-1937.75, 849.64, 410.36) mm, rotated rx -89.89 ry 0.49 rz -179.51 deg; joints [-25.805, 39.339, 0.414, -72.391, 33.595, -44.539, -170]
  MoveL 240 to (-1937.75, 849.7, 440.36) mm, rotated rx -89.89 ry 0.48 rz -179.52 deg; joints [-25.822, 38.483, 0.372, -70.411, 31.663, -45.097, -170]
  MoveL 241 to (-1937.75, 849.75, 470.36) mm, rotated rx -89.89 ry 0.48 rz -179.53 deg; joints [-25.842, 37.642, 0.302, -68.267, 29.629, -45.757, -170]
  MoveL 242 to (-1937.75, 849.81, 500.36) mm, rotated rx -89.89 ry 0.47 rz -179.53 deg; joints [-25.866, 36.816, 0.201, -65.925, 27.474, -46.542, -170]
  MoveL 243 to (-1937.75, 849.86, 530.36) mm, rotated rx -89.88 ry 0.46 rz -179.54 deg; joints [-25.894, 36.006, 0.07, -63.335, 25.166, -47.482, -170]
  MoveL 244 to (-1937.75, 849.91, 554.46) mm, rotated rx -89.88 ry 0.46 rz -179.54 deg; joints [-25.921, 35.367, -0.058, -61.025, 23.174, -48.382, -170]
  MoveL 245 to (-1937.75, 849.96, 584.46) mm, rotated rx -89.9 ry 0.45 rz -179.56 deg; joints [-25.961, 34.582, -0.252, -57.675, 20.395, -49.775, -170]
  MoveL 246 to (-1937.75, 850.01, 614.46) mm, rotated rx -89.91 ry 0.44 rz -179.57 deg; joints [-26.013, 33.815, -0.483, -53.682, 17.228, -51.569, -170]
  MoveL 247 to (-1937.75, 850.06, 644.46) mm, rotated rx -89.93 ry 0.42 rz -179.58 deg; joints [-26.087, 33.064, -0.759, -48.595, 13.394, -54.041, -170]
  MoveL 248 to (-1937.75, 850.09, 662.91) mm, rotated rx -89.93 ry 0.42 rz -179.59 deg; joints [-26.153, 32.611, -0.959, -44.405, 10.383, -56.211, -170]
  MoveL 249 to (-1937.75, 850.1, 692.91) mm, rotated rx -89.97 ry 20.4 rz -179.59 deg; joints [-25.413, 34.856, -0.195, -90.022, 57.282, -31.269, -170]
  MoveL 250 to (-1937.75, 850.1, 722.91) mm, rotated rx -90.02 ry 20.38 rz -179.62 deg; joints [-25.414, 34.092, -0.38, -88.573, 55.554, -31.284, -170]
  MoveL 251 to (-1937.75, 850.1, 752.91) mm, rotated rx -90.06 ry 20.37 rz -179.65 deg; joints [-25.417, 33.346, -0.593, -87.079, 53.796, -31.333, -170]
  MoveL 252 to (-1937.75, 850.1, 771.36) mm, rotated rx -90.08 ry 20.36 rz -179.67 deg; joints [-25.418, 32.896, -0.738, -86.137, 52.699, -31.381, -170]
  MoveL 253 to (-1937.75, 849.97, 801.36) mm, rotated rx -92.77 ry 22.38 rz 179.05 deg; joints [-25.207, 31.933, -1.211, -82.424, 50.699, -29.873, -170]
  MoveL 254 to (-1937.75, 849.83, 831.36) mm, rotated rx -95.32 ry 18.12 rz 178.19 deg; joints [-25.327, 30.092, -1.895, -69.323, 36.37, -32.97, -170]
  MoveL 255 to (-1937.75, 849.69, 861.36) mm, rotated rx -97.87 ry 16.65 rz 177.32 deg; joints [-25.424, 28.806, -2.796, -56.793, 25.497, -36.599, -170]
  MoveL 256 to (-1937.75, 849.61, 879.82) mm, rotated rx -99.44 ry 16.1 rz 176.79 deg; joints [-25.542, 28.121, -3.45, -46.824, 17.915, -40.416, -170]
  MoveL 257 to (-1937.75, 849.61, 879.82) mm, rotated rx -99.44 ry 16.1 rz 176.79 deg; joints [-25.542, 28.121, -3.45, -46.824, 17.915, -40.416, -170]
  MoveL 258 to (-1937.75, 840.64, 908.44) mm, rotated rx -99.35 ry 16.95 rz 176.82 deg; joints [-25.739, 27.906, -4.079, -47.048, 17.949, -39.762, -170]
  MoveL 259 to (-1937.75, 830.31, 941.39) mm, rotated rx -99.26 ry 17.96 rz 176.85 deg; joints [-25.96, 27.686, -4.828, -47.373, 18.064, -38.963, -170]
  MoveL 260 to (-1937.75, 821.74, 970.15) mm, rotated rx -105.49 ry 37.99 rz 170.12 deg; joints [-24.576, 29.536, -5.647, -70.942, 52.152, -22.559, -170]
  MoveL 261 to (-1937.75, 811.88, 1003.24) mm, rotated rx -110.4 ry 37.75 rz 167.06 deg; joints [-24.796, 28.511, -7.141, -60.377, 43.492, -23.298, -170]
  MoveL 262 to (-1937.75, 803.91, 1032.16) mm, rotated rx -109.88 ry 39.18 rz 167.37 deg; joints [-24.944, 28.485, -7.721, -62.182, 45.192, -22.374, -170]
  MoveL 263 to (-1937.75, 798.76, 1050.87) mm, rotated rx -109.55 ry 40.17 rz 167.57 deg; joints [-25.035, 28.487, -8.113, -63.366, 46.374, -21.769, -170]
  Set speed (1000.0 mm/s)
  MoveL 264 to (-1937.75, 798.76, 1050.87) mm, rotated rx -109.55 ry 40.17 rz 167.57 deg; joints [-25.035, 28.487, -8.113, -63.366, 46.374, -21.769, -170]
  MoveL 265 to (-1938.54, 895.43, 1076.44) mm, rotated rx -109.55 ry 40.17 rz 167.57 deg; joints [-22.959, 25.504, -4.981, -61.386, 46.769, -24.193, -170]
  Set speed (1000.0 mm/s)
  MoveL 266 to (-2018.52, 892.55, 1084.66) mm, rotated rx -110.44 ry 39.9 rz 167.02 deg; joints [-24.417, 22.763, -1.795, -62.483, 46.476, -22.232, -170]
  MoveL 267 to (-2017.75, 796.21, 1057.87) mm, rotated rx -110.44 ry 39.9 rz 167.02 deg; joints [-26.5, 25.824, -4.863, -64.872, 46.45, -19.677, -170]
  MoveL 268 to (-2017.75, 796.21, 1057.87) mm, rotated rx -110.44 ry 39.9 rz 167.02 deg; joints [-26.5, 25.824, -4.863, -64.872, 46.45, -19.677, -170]
  Set speed (50.0 mm/s)
  MoveL 269 to (-2017.75, 801.6, 1039.29) mm, rotated rx -110.46 ry 39.83 rz 167.01 deg; joints [-26.372, 25.978, -4.342, -65.932, 47.621, -19.474, -170]
  MoveL 270 to (-2017.75, 809.95, 1010.47) mm, rotated rx -111.29 ry 37.47 rz 166.51 deg; joints [-26.244, 25.838, -3.894, -61.866, 43.525, -21.217, -170]
  MoveL 271 to (-2017.75, 820.22, 977.55) mm, rotated rx -103.38 ry 18.44 rz 175.46 deg; joints [-27.962, 24.375, -3.19, -30.396, 5.105, -43.823, -170]
  MoveL 272 to (-2017.75, 829.16, 948.91) mm, rotated rx -99.61 ry 17.86 rz 176.73 deg; joints [-27.381, 25.14, -1.517, -53.742, 21.201, -34.616, -170]
  MoveL 273 to (-2017.75, 839.86, 916.11) mm, rotated rx -99.68 ry 16.86 rz 176.7 deg; joints [-27.146, 25.357, -0.747, -53.531, 21.178, -35.391, -170]
  MoveL 274 to (-2017.75, 849.17, 887.6) mm, rotated rx -99.75 ry 16.02 rz 176.68 deg; joints [-26.939, 25.569, -0.099, -53.378, 21.204, -36.042, -170]
  MoveL 275 to (-2017.75, 849.24, 868.13) mm, rotated rx -98.05 ry 16.59 rz 177.26 deg; joints [-26.849, 26.315, 0.591, -62.468, 28.478, -33.062, -170]
  MoveL 276 to (-2017.75, 849.36, 838.13) mm, rotated rx -95.42 ry 18.04 rz 178.15 deg; joints [-26.783, 27.642, 1.499, -73.878, 38.879, -30.385, -170]
  MoveL 277 to (-2017.75, 849.48, 808.13) mm, rotated rx -92.8 ry 22.28 rz 179.04 deg; joints [-26.684, 29.531, 2.201, -86.163, 52.938, -28.076, -170]
  MoveL 278 to (-2017.75, 849.59, 778.13) mm, rotated rx -90.04 ry 20.36 rz -179.65 deg; joints [-26.908, 30.564, 2.673, -90.103, 55.305, -29.7, -170]
  MoveL 279 to (-2017.75, 849.58, 758.66) mm, rotated rx -90.02 ry 20.37 rz -179.64 deg; joints [-26.907, 31.052, 2.827, -91.062, 56.462, -29.708, -170]
  MoveL 280 to (-2017.75, 849.56, 728.66) mm, rotated rx -89.98 ry 0.39 rz -179.61 deg; joints [-27.672, 28.854, 1.867, -44.977, 8.865, -54.909, -170]
  MoveL 281 to (-2017.75, 849.54, 698.66) mm, rotated rx -89.94 ry 0.4 rz -179.6 deg; joints [-27.559, 29.582, 2.262, -52.251, 14.115, -51.187, -170]
  MoveL 282 to (-2017.75, 849.52, 668.66) mm, rotated rx -89.9 ry 0.42 rz -179.58 deg; joints [-27.491, 30.328, 2.59, -57.205, 17.935, -48.884, -170]
  MoveL 283 to (-2017.75, 849.48, 649.19) mm, rotated rx -89.9 ry 0.43 rz -179.58 deg; joints [-27.459, 30.819, 2.773, -59.768, 20.007, -47.771, -170]
  MoveL 284 to (-2017.75, 849.41, 619.19) mm, rotated rx -89.88 ry 0.44 rz -179.56 deg; joints [-27.419, 31.591, 3.025, -63.184, 22.876, -46.39, -170]
  MoveL 285 to (-2017.75, 849.35, 589.19) mm, rotated rx -89.87 ry 0.45 rz -179.55 deg; joints [-27.388, 32.38, 3.241, -66.144, 25.468, -45.294, -170]
  MoveL 286 to (-2017.75, 849.28, 559.19) mm, rotated rx -89.86 ry 0.46 rz -179.54 deg; joints [-27.363, 33.187, 3.425, -68.773, 27.86, -44.407, -170]
  MoveL 287 to (-2017.75, 849.22, 531.21) mm, rotated rx -89.86 ry 0.47 rz -179.54 deg; joints [-27.342, 33.95, 3.566, -70.941, 29.908, -43.736, -170]
  MoveL 288 to (-2017.75, 849.16, 501.21) mm, rotated rx -89.86 ry 0.47 rz -179.53 deg; joints [-27.324, 34.784, 3.688, -73.079, 31.988, -43.134, -170]
  MoveL 289 to (-2017.75, 849.09, 471.21) mm, rotated rx -89.87 ry 0.48 rz -179.52 deg; joints [-27.308, 35.635, 3.781, -75.056, 33.968, -42.633, -170]
  MoveL 290 to (-2017.75, 849.03, 441.21) mm, rotated rx -89.87 ry 0.48 rz -179.52 deg; joints [-27.294, 36.501, 3.846, -76.901, 35.863, -42.216, -170]
  MoveL 291 to (-2017.75, 848.96, 411.21) mm, rotated rx -89.87 ry 0.49 rz -179.51 deg; joints [-27.282, 37.382, 3.882, -78.631, 37.685, -41.869, -170]
  MoveL 292 to (-2017.75, 848.9, 381.21) mm, rotated rx -89.88 ry 0.5 rz -179.51 deg; joints [-27.272, 38.278, 3.891, -80.262, 39.441, -41.583, -170]
  MoveL 293 to (-2017.75, 848.84, 351.21) mm, rotated rx -89.88 ry 0.5 rz -179.5 deg; joints [-27.263, 39.188, 3.873, -81.808, 41.139, -41.35, -170]
  MoveL 294 to (-2017.75, 848.77, 321.21) mm, rotated rx -89.88 ry 0.51 rz -179.49 deg; joints [-27.255, 40.112, 3.827, -83.276, 42.783, -41.163, -170]
  MoveL 295 to (-2017.75, 848.71, 291.21) mm, rotated rx -89.89 ry 0.51 rz -179.49 deg; joints [-27.249, 41.05, 3.753, -84.676, 44.378, -41.016, -170]
  MoveL 296 to (-2017.75, 848.64, 261.21) mm, rotated rx -89.89 ry 0.52 rz -179.48 deg; joints [-27.243, 42.001, 3.654, -86.014, 45.927, -40.905, -170]
  MoveL 297 to (-2017.75, 848.58, 231.21) mm, rotated rx -89.89 ry 0.53 rz -179.48 deg; joints [-27.238, 42.965, 3.527, -87.296, 47.434, -40.825, -170]
  MoveL 298 to (-2017.75, 848.52, 201.21) mm, rotated rx -89.9 ry 0.53 rz -179.47 deg; joints [-27.233, 43.941, 3.373, -88.526, 48.899, -40.774, -170]
  MoveL 299 to (-2017.75, 848.5, 193.21) mm, rotated rx -89.9 ry 0.53 rz -179.47 deg; joints [-27.232, 44.203, 3.328, -88.84, 49.279, -40.768, -170]
  Set speed (1000.0 mm/s)
  MoveL 300 to (-2017.75, 848.5, 193.21) mm, rotated rx -89.9 ry 0.53 rz -179.47 deg; joints [-27.232, 44.203, 3.328, -88.84, 49.279, -40.768, -170]
  MoveL 301 to (-2018.67, 948.49, 193.03) mm, rotated rx -89.9 ry 0.53 rz -179.47 deg; joints [-24.993, 42.229, 6.952, -87.511, 51.213, -42.753, -170]
  Set speed (1000.0 mm/s)
  MoveL 302 to (-2098.68, 947.75, 193.86) mm, rotated rx -89.89 ry 0.54 rz -179.46 deg; joints [-26.586, 40.53, 10.242, -92.377, 54.643, -41.382, -170]
  MoveL 303 to (-2097.75, 847.76, 194.06) mm, rotated rx -89.89 ry 0.54 rz -179.46 deg; joints [-28.84, 42.519, 6.596, -93.821, 52.814, -39.352, -170]
  MoveL 304 to (-2097.75, 847.76, 194.06) mm, rotated rx -89.89 ry 0.54 rz -179.46 deg; joints [-28.84, 42.519, 6.596, -93.821, 52.814, -39.352, -170]
  Set speed (50.0 mm/s)
  MoveL 305 to (-2097.75, 847.78, 202.06) mm, rotated rx -89.89 ry 0.54 rz -179.46 deg; joints [-28.841, 42.25, 6.643, -93.523, 52.436, -39.332, -170]
  MoveL 306 to (-2097.75, 847.85, 232.06) mm, rotated rx -89.88 ry 0.53 rz -179.47 deg; joints [-28.841, 41.248, 6.797, -92.345, 50.971, -39.298, -170]
  MoveL 307 to (-2097.75, 847.92, 262.06) mm, rotated rx -89.88 ry 0.52 rz -179.48 deg; joints [-28.844, 40.258, 6.927, -91.144, 49.482, -39.272, -170]
  MoveL 308 to (-2097.75, 848, 292.06) mm, rotated rx -89.87 ry 0.52 rz -179.49 deg; joints [-28.847, 39.28, 7.03, -89.897, 47.956, -39.271, -170]
  MoveL 309 to (-2097.75, 848.07, 322.06) mm, rotated rx -89.87 ry 0.51 rz -179.49 deg; joints [-28.851, 38.316, 7.106, -88.601, 46.39, -39.298, -170]
  MoveL 310 to (-2097.75, 848.14, 352.06) mm, rotated rx -89.86 ry 0.5 rz -179.5 deg; joints [-28.856, 37.365, 7.156, -87.251, 44.784, -39.355, -170]
  MoveL 311 to (-2097.75, 848.21, 382.06) mm, rotated rx -89.86 ry 0.5 rz -179.5 deg; joints [-28.861, 36.428, 7.178, -85.842, 43.133, -39.448, -170]
  MoveL 312 to (-2097.75, 848.29, 412.06) mm, rotated rx -89.85 ry 0.49 rz -179.51 deg; joints [-28.868, 35.506, 7.173, -84.367, 41.435, -39.58, -170]
  MoveL 313 to (-2097.75, 848.36, 442.06) mm, rotated rx -89.85 ry 0.49 rz -179.52 deg; joints [-28.876, 34.599, 7.141, -82.817, 39.685, -39.758, -170]
  MoveL 314 to (-2097.75, 848.43, 472.06) mm, rotated rx -89.85 ry 0.48 rz -179.52 deg; joints [-28.885, 33.708, 7.081, -81.184, 37.879, -39.988, -170]
  MoveL 315 to (-2097.75, 848.5, 502.06) mm, rotated rx -89.84 ry 0.47 rz -179.53 deg; joints [-28.895, 32.832, 6.994, -79.455, 36.01, -40.277, -170]
  MoveL 316 to (-2097.75, 848.58, 532.06) mm, rotated rx -89.84 ry 0.47 rz -179.53 deg; joints [-28.907, 31.972, 6.878, -77.615, 34.068, -40.636, -170]
  MoveL 317 to (-2097.75, 848.65, 563.91) mm, rotated rx -89.83 ry 0.46 rz -179.54 deg; joints [-28.923, 31.078, 6.723, -75.518, 31.916, -41.109, -170]
  MoveL 318 to (-2097.75, 848.73, 593.91) mm, rotated rx -89.84 ry 0.45 rz -179.55 deg; joints [-28.939, 30.249, 6.545, -73.321, 29.74, -41.67, -170]
  MoveL 319 to (-2097.75, 848.81, 623.91) mm, rotated rx -89.86 ry 0.44 rz -179.56 deg; joints [-28.958, 29.438, 6.336, -70.92, 27.439, -42.36, -170]
  MoveL 320 to (-2097.75, 848.89, 653.91) mm, rotated rx -89.87 ry 0.43 rz -179.57 deg; joints [-28.982, 28.644, 6.096, -68.258, 24.979, -43.216, -170]
  MoveL 321 to (-2097.75, 848.95, 674.4) mm, rotated rx -89.88 ry 0.42 rz -179.58 deg; joints [-29.002, 28.114, 5.912, -66.249, 23.183, -43.921, -170]
  MoveL 322 to (-2097.75, 848.99, 704.4) mm, rotated rx -89.91 ry 0.41 rz -179.6 deg; joints [-29.039, 27.347, 5.608, -62.83, 20.246, -45.219, -170]
  MoveL 323 to (-2097.75, 849.02, 734.4) mm, rotated rx -89.95 ry 0.39 rz -179.61 deg; joints [-29.088, 26.601, 5.263, -58.718, 16.89, -46.948, -170]
  MoveL 324 to (-2097.75, 849.06, 764.4) mm, rotated rx -89.98 ry 0.38 rz -179.63 deg; joints [-29.161, 25.874, 4.867, -53.374, 12.78, -49.437, -170]
  MoveL 325 to (-2097.75, 849.08, 784.89) mm, rotated rx -90.01 ry 0.37 rz -179.64 deg; joints [-29.241, 25.389, 4.553, -48.173, 9.013, -52.083, -170]
  MoveL 326 to (-2097.75, 848.99, 814.89) mm, rotated rx -92.84 ry 22.17 rz 179.02 deg; joints [-28.259, 27.194, 5.435, -89.802, 55.025, -26.318, -170]
  MoveL 327 to (-2097.75, 848.89, 844.89) mm, rotated rx -95.53 ry 17.96 rz 178.11 deg; joints [-28.339, 25.256, 4.713, -78.221, 41.185, -27.911, -170]
  MoveL 328 to (-2097.75, 848.79, 874.89) mm, rotated rx -98.24 ry 16.52 rz 177.19 deg; joints [-28.379, 23.888, 3.795, -67.686, 31.118, -29.789, -170]
  MoveL 329 to (-2097.75, 848.73, 895.37) mm, rotated rx -100.08 ry 15.94 rz 176.57 deg; joints [-28.446, 23.08, 3.063, -59.153, 23.948, -32.115, -170]
  MoveL 330 to (-2097.75, 848.73, 895.37) mm, rotated rx -100.08 ry 15.94 rz 176.57 deg; joints [-28.446, 23.08, 3.063, -59.153, 23.948, -32.115, -170]
  MoveL 331 to (-2097.75, 839.07, 923.78) mm, rotated rx -100.02 ry 16.78 rz 176.59 deg; joints [-28.664, 22.874, 2.395, -59.279, 23.892, -31.44, -170]
  MoveL 332 to (-2097.75, 827.93, 956.54) mm, rotated rx -99.96 ry 17.77 rz 176.61 deg; joints [-28.911, 22.662, 1.6, -59.439, 23.865, -30.647, -170]
  MoveL 333 to (-2097.75, 818.63, 985.06) mm, rotated rx -103.93 ry 18.32 rz 175.28 deg; joints [-29.382, 21.874, -0.093, -41.445, 10.78, -36.206, -170]
  MoveL 334 to (-2097.75, 807.9, 1017.96) mm, rotated rx -112.2 ry 37.2 rz 165.94 deg; joints [-27.785, 23.239, -0.857, -63.271, 43.368, -19.079, -170]
  MoveL 335 to (-2097.75, 799.15, 1046.65) mm, rotated rx -111.71 ry 38.58 rz 166.24 deg; joints [-27.956, 23.216, -1.453, -64.924, 44.94, -18.195, -170]
  MoveL 336 to (-2097.75, 793.47, 1065.33) mm, rotated rx -111.4 ry 39.53 rz 166.43 deg; joints [-28.063, 23.218, -1.854, -66.002, 46.028, -17.618, -170]
  Set speed (1000.0 mm/s)
  MoveL 337 to (-2097.75, 793.47, 1065.33) mm, rotated rx -111.4 ry 39.53 rz 166.43 deg; joints [-28.063, 23.218, -1.854, -66.002, 46.028, -17.618, -170]
  MoveL 338 to (-2098.47, 889.42, 1093.47) mm, rotated rx -111.4 ry 39.53 rz 166.43 deg; joints [-25.98, 20.067, 1.151, -63.175, 45.656, -20.311, -170]
  Set speed (1000.0 mm/s)
  MoveL 339 to (-2178.49, 886.05, 1102.66) mm, rotated rx -112.35 ry 39.32 rz 165.84 deg; joints [-27.647, 17.456, 3.914, -64.127, 44.978, -18.171, -170]
  MoveL 340 to (-2177.75, 790.48, 1073.24) mm, rotated rx -112.35 ry 39.32 rz 165.84 deg; joints [-29.723, 20.707, 0.959, -67.381, 45.756, -15.356, -170]
  MoveL 341 to (-2177.75, 790.48, 1073.24) mm, rotated rx -112.35 ry 39.32 rz 165.84 deg; joints [-29.723, 20.707, 0.959, -67.381, 45.756, -15.356, -170]
  Set speed (50.0 mm/s)
  MoveL 342 to (-2177.75, 796.55, 1054.26) mm, rotated rx -112.37 ry 39.26 rz 165.83 deg; joints [-29.578, 20.851, 1.53, -68.498, 47.027, -15.177, -170]
  MoveL 343 to (-2177.75, 805.69, 1025.69) mm, rotated rx -113.14 ry 36.95 rz 165.37 deg; joints [-29.426, 20.709, 1.976, -64.616, 43.028, -16.863, -170]
  MoveL 344 to (-2177.75, 816.95, 992.69) mm, rotated rx -104.49 ry 18.22 rz 175.09 deg; joints [-30.974, 19.446, 2.79, -49.235, 14.364, -30.524, -170]
  MoveL 345 to (-2177.75, 826.64, 964.3) mm, rotated rx -100.33 ry 17.69 rz 176.49 deg; joints [-30.552, 20.251, 4.532, -64.761, 26.236, -26.875, -170]
  MoveL 346 to (-2177.75, 838.27, 931.43) mm, rotated rx -100.38 ry 16.7 rz 176.47 deg; joints [-30.292, 20.453, 5.358, -64.616, 26.285, -27.71, -170]
  MoveL 347 to (-2177.75, 848.29, 903.15) mm, rotated rx -100.42 ry 15.86 rz 176.45 deg; joints [-30.064, 20.65, 6.048, -64.491, 26.353, -28.424, -170]
  MoveL 348 to (-2177.75, 848.34, 881.65) mm, rotated rx -98.43 ry 16.46 rz 177.13 deg; joints [-30.017, 21.522, 6.825, -72.625, 33.524, -26.671, -170]
  MoveL 349 to (-2177.75, 848.42, 851.65) mm, rotated rx -95.65 ry 17.88 rz 178.07 deg; joints [-30.001, 22.933, 7.757, -82.438, 43.341, -25.497, -170]
  MoveL 350 to (-2177.75, 848.5, 821.65) mm, rotated rx -92.67 ry 2.07 rz 180 deg; joints [-30.801, 22.121, 7.035, -53.396, 11.005, -45.105, -170]
  MoveL 351 to (-2177.75, 848.58, 791.65) mm, rotated rx -89.97 ry 0.37 rz -179.63 deg; joints [-30.768, 23.146, 7.771, -61.643, 16.755, -44.218, -170]
  MoveL 352 to (-2177.75, 848.54, 770.15) mm, rotated rx -89.95 ry 0.38 rz -179.62 deg; joints [-30.734, 23.667, 8.059, -64.62, 19.213, -42.997, -170]
  MoveL 353 to (-2177.75, 848.48, 740.15) mm, rotated rx -89.91 ry 0.4 rz -179.61 deg; joints [-30.697, 24.413, 8.425, -68.138, 22.256, -41.689, -170]
  MoveL 354 to (-2177.75, 848.43, 710.15) mm, rotated rx -89.88 ry 0.41 rz -179.59 deg; joints [-30.67, 25.179, 8.753, -71.157, 24.996, -40.692, -170]
  MoveL 355 to (-2177.75, 848.38, 680.15) mm, rotated rx -89.85 ry 0.42 rz -179.58 deg; joints [-30.648, 25.965, 9.047, -73.827, 27.524, -39.916, -170]
  MoveL 356 to (-2177.75, 848.31, 658.64) mm, rotated rx -89.84 ry 0.43 rz -179.57 deg; joints [-30.636, 26.537, 9.234, -75.53, 29.195, -39.47, -170]
  MoveL 357 to (-2177.75, 848.22, 628.64) mm, rotated rx -89.83 ry 0.44 rz -179.56 deg; joints [-30.621, 27.352, 9.469, -77.731, 31.42, -38.958, -170]
  MoveL 358 to (-2177.75, 848.12, 598.64) mm, rotated rx -89.82 ry 0.45 rz -179.55 deg; joints [-30.61, 28.186, 9.674, -79.765, 33.54, -38.553, -170]
  MoveL 359 to (-2177.75, 848.03, 568.64) mm, rotated rx -89.81 ry 0.46 rz -179.54 deg; joints [-30.6, 29.037, 9.849, -81.66, 35.574, -38.236, -170]
  MoveL 360 to (-2177.75, 847.93, 532.9) mm, rotated rx -89.81 ry 0.47 rz -179.53 deg; joints [-30.589, 30.07, 10.018, -83.717, 37.855, -37.959, -170]
  MoveL 361 to (-2177.75, 847.85, 502.9) mm, rotated rx -89.82 ry 0.48 rz -179.53 deg; joints [-30.582, 30.955, 10.129, -85.341, 39.703, -37.792, -170]
  MoveL 362 to (-2177.75, 847.77, 472.9) mm, rotated rx -89.82 ry 0.48 rz -179.52 deg; joints [-30.575, 31.857, 10.212, -86.885, 41.496, -37.674, -170]
  MoveL 363 to (-2177.75, 847.69, 442.9) mm, rotated rx -89.83 ry 0.49 rz -179.51 deg; joints [-30.57, 32.775, 10.268, -88.358, 43.241, -37.602, -170]
  MoveL 364 to (-2177.75, 847.61, 412.9) mm, rotated rx -89.84 ry 0.49 rz -179.51 deg; joints [-30.566, 33.709, 10.296, -89.768, 44.94, -37.568, -170]
  MoveL 365 to (-2177.75, 847.53, 382.9) mm, rotated rx -89.84 ry 0.5 rz -179.5 deg; joints [-30.562, 34.658, 10.298, -91.122, 46.598, -37.568, -170]
  MoveL 366 to (-2177.75, 847.45, 352.9) mm, rotated rx -89.85 ry 0.51 rz -179.5 deg; joints [-30.56, 35.622, 10.272, -92.424, 48.216, -37.599, -170]
  MoveL 367 to (-2177.75, 847.36, 322.9) mm, rotated rx -89.85 ry 0.51 rz -179.49 deg; joints [-30.557, 36.6, 10.219, -93.68, 49.797, -37.657, -170]
  MoveL 368 to (-2177.75, 847.28, 292.9) mm, rotated rx -89.86 ry 0.52 rz -179.49 deg; joints [-30.556, 37.592, 10.139, -94.894, 51.344, -37.739, -170]
  MoveL 369 to (-2177.75, 847.2, 262.9) mm, rotated rx -89.86 ry 0.52 rz -179.48 deg; joints [-30.555, 38.597, 10.033, -96.068, 52.856, -37.843, -170]
  MoveL 370 to (-2177.75, 847.12, 232.9) mm, rotated rx -89.87 ry 0.53 rz -179.47 deg; joints [-30.554, 39.615, 9.9, -97.205, 54.335, -37.966, -170]
  MoveL 371 to (-2177.75, 847.04, 202.9) mm, rotated rx -89.87 ry 0.53 rz -179.47 deg; joints [-30.554, 40.645, 9.741, -98.307, 55.782, -38.107, -170]
  MoveL 372 to (-2177.75, 847.02, 194.9) mm, rotated rx -89.87 ry 0.53 rz -179.47 deg; joints [-30.554, 40.922, 9.694, -98.591, 56.161, -38.15, -170]
  Set speed (1000.0 mm/s)
  MoveL 373 to (-2177.75, 847.02, 194.9) mm, rotated rx -89.87 ry 0.53 rz -179.47 deg; joints [-30.554, 40.922, 9.694, -98.591, 56.161, -38.15, -170]
  MoveL 374 to (-2178.67, 947.01, 194.68) mm, rotated rx -89.87 ry 0.53 rz -179.47 deg; joints [-28.29, 38.913, 13.37, -97.067, 57.905, -40.211, -170]
  Set speed (1000.0 mm/s)
  MoveL 375 to (-2258.68, 946.27, 195.52) mm, rotated rx -89.86 ry 0.54 rz -179.46 deg; joints [-30.123, 37.37, 16.349, -101.71, 61.065, -39.155, -170]
  MoveL 376 to (-2257.75, 846.28, 195.75) mm, rotated rx -89.86 ry 0.54 rz -179.46 deg; joints [-32.386, 39.405, 12.632, -103.285, 59.392, -37.073, -170]
  MoveL 377 to (-2257.75, 846.28, 195.75) mm, rotated rx -89.86 ry 0.54 rz -179.46 deg; joints [-32.386, 39.405, 12.632, -103.285, 59.392, -37.073, -170]
  Set speed (50.0 mm/s)
  MoveL 378 to (-2257.75, 846.3, 203.75) mm, rotated rx -89.86 ry 0.54 rz -179.46 deg; joints [-32.386, 39.121, 12.68, -103.012, 59.014, -37.007, -170]
  MoveL 379 to (-2257.75, 846.39, 233.75) mm, rotated rx -89.85 ry 0.53 rz -179.47 deg; joints [-32.383, 38.064, 12.841, -101.941, 57.56, -36.792, -170]
  MoveL 380 to (-2257.75, 846.48, 263.75) mm, rotated rx -89.85 ry 0.52 rz -179.48 deg; joints [-32.381, 37.017, 12.977, -100.857, 56.086, -36.576, -170]
  MoveL 381 to (-2257.75, 846.57, 293.75) mm, rotated rx -89.84 ry 0.52 rz -179.48 deg; joints [-32.38, 35.984, 13.087, -99.743, 54.583, -36.376, -170]
  MoveL 382 to (-2257.75, 846.66, 323.75) mm, rotated rx -89.83 ry 0.51 rz -179.49 deg; joints [-32.38, 34.963, 13.17, -98.598, 53.05, -36.193, -170]
  MoveL 383 to (-2257.75, 846.75, 353.75) mm, rotated rx -89.83 ry 0.51 rz -179.5 deg; joints [-32.379, 33.957, 13.226, -97.419, 51.487, -36.028, -170]
  MoveL 384 to (-2257.75, 846.84, 383.75) mm, rotated rx -89.82 ry 0.5 rz -179.5 deg; joints [-32.38, 32.965, 13.255, -96.204, 49.892, -35.884, -170]
  MoveL 385 to (-2257.75, 846.93, 413.75) mm, rotated rx -89.82 ry 0.5 rz -179.51 deg; joints [-32.381, 31.988, 13.257, -94.949, 48.264, -35.763, -170]
  MoveL 386 to (-2257.75, 847.02, 443.75) mm, rotated rx -89.81 ry 0.49 rz -179.51 deg; joints [-32.382, 31.027, 13.232, -93.651, 46.602, -35.669, -170]
  MoveL 387 to (-2257.75, 847.11, 473.75) mm, rotated rx -89.81 ry 0.48 rz -179.52 deg; joints [-32.384, 30.081, 13.18, -92.306, 44.904, -35.604, -170]
  MoveL 388 to (-2257.75, 847.19, 503.75) mm, rotated rx -89.8 ry 0.48 rz -179.52 deg; joints [-32.387, 29.153, 13.1, -90.908, 43.167, -35.572, -170]
  MoveL 389 to (-2257.75, 847.28, 533.75) mm, rotated rx -89.79 ry 0.47 rz -179.53 deg; joints [-32.391, 28.241, 12.993, -89.452, 41.388, -35.578, -170]
  MoveL 390 to (-2257.75, 847.4, 573.37) mm, rotated rx -89.79 ry 0.47 rz -179.54 deg; joints [-32.398, 27.064, 12.809, -87.425, 38.967, -35.652, -170]
  MoveL 391 to (-2257.75, 847.51, 603.37) mm, rotated rx -89.79 ry 0.46 rz -179.55 deg; joints [-32.403, 26.189, 12.635, -85.758, 37.035, -35.769, -170]
  MoveL 392 to (-2257.75, 847.62, 633.37) mm, rotated rx -89.8 ry 0.45 rz -179.56 deg; joints [-32.409, 25.333, 12.433, -83.994, 35.041, -35.949, -170]
  MoveL 393 to (-2257.75, 847.72, 663.37) mm, rotated rx -89.81 ry 0.43 rz -179.57 deg; joints [-32.417, 24.497, 12.202, -82.117, 32.974, -36.202, -170]
  MoveL 394 to (-2257.75, 847.8, 685.89) mm, rotated rx -89.82 ry 0.43 rz -179.57 deg; joints [-32.424, 23.882, 12.009, -80.62, 31.369, -36.449, -170]
  MoveL 395 to (-2257.75, 847.87, 715.89) mm, rotated rx -89.85 ry 0.41 rz -179.59 deg; joints [-32.436, 23.075, 11.721, -78.427, 29.088, -36.873, -170]
  MoveL 396 to (-2257.75, 847.94, 745.89) mm, rotated rx -89.88 ry 0.4 rz -179.6 deg; joints [-32.451, 22.29, 11.401, -76.026, 26.681, -37.43, -170]
  MoveL 397 to (-2257.75, 848.01, 775.89) mm, rotated rx -89.91 ry 0.38 rz -179.62 deg; joints [-32.471, 21.526, 11.048, -73.356, 24.11, -38.157, -170]
  MoveL 398 to (-2257.75, 848.06, 798.41) mm, rotated rx -89.93 ry 0.37 rz -179.63 deg; joints [-32.489, 20.966, 10.76, -71.12, 22.039, -38.85, -170]
  MoveL 399 to (-2257.75, 848.01, 828.41) mm, rotated rx -92.71 ry 1.95 rz 180 deg; joints [-32.469, 19.884, 10.033, -64.813, 17.224, -38.316, -170]
  MoveL 400 to (-2257.75, 847.95, 858.41) mm, rotated rx -95.77 ry 17.8 rz 178.03 deg; joints [-31.774, 20.67, 10.637, -86.595, 45.391, -23.104, -170]
  MoveL 401 to (-2257.75, 847.89, 888.41) mm, rotated rx -98.64 ry 16.4 rz 177.06 deg; joints [-31.768, 19.217, 9.689, -77.409, 35.771, -23.632, -170]
  MoveL 402 to (-2257.75, 847.85, 910.93) mm, rotated rx -100.78 ry 15.78 rz 176.33 deg; joints [-31.796, 18.28, 8.863, -69.595, 28.542, -24.841, -170]
  MoveL 403 to (-2257.75, 847.85, 910.93) mm, rotated rx -100.78 ry 15.78 rz 176.33 deg; joints [-31.796, 18.28, 8.863, -69.595, 28.542, -24.841, -170]
  MoveL 404 to (-2257.75, 837.46, 939.08) mm, rotated rx -100.75 ry 16.62 rz 176.35 deg; joints [-32.034, 18.095, 8.15, -69.734, 28.477, -24.082, -170]
  MoveL 405 to (-2257.75, 825.25, 972.18) mm, rotated rx -100.71 ry 17.62 rz 176.36 deg; joints [-32.308, 17.906, 7.286, -69.888, 28.422, -23.189, -170]
  MoveL 406 to (-2257.75, 815.17, 1000.43) mm, rotated rx -105.06 ry 18.12 rz 174.9 deg; joints [-32.696, 17.089, 5.487, -56.077, 17.303, -25.391, -170]
  MoveL 407 to (-2257.75, 803.32, 1033.66) mm, rotated rx -114.11 ry 36.7 rz 164.78 deg; joints [-31.172, 18.248, 4.612, -65.933, 42.52, -14.546, -170]
  MoveL 408 to (-2257.75, 793.77, 1062.1) mm, rotated rx -113.66 ry 38.05 rz 165.05 deg; joints [-31.365, 18.242, 3.987, -67.459, 43.997, -13.662, -170]
  MoveL 409 to (-2257.75, 787.22, 1081.61) mm, rotated rx -113.37 ry 39.02 rz 165.22 deg; joints [-31.494, 18.254, 3.545, -68.499, 45.067, -13.059, -170]
  Set speed (1000.0 mm/s)
  MoveL 410 to (-2257.75, 787.22, 1081.61) mm, rotated rx -113.37 ry 39.02 rz 165.22 deg; joints [-31.494, 18.254, 3.545, -68.499, 45.067, -13.059, -170]
  MoveL 411 to (-2258.48, 882.35, 1112.44) mm, rotated rx -113.37 ry 39.02 rz 165.22 deg; joints [-29.434, 14.894, 6.448, -64.781, 43.845, -16.006, -170]
  Set speed (1000.0 mm/s)
  MoveL 412 to (-2338.51, 878.31, 1122.67) mm, rotated rx -114.42 ry 38.8 rz 164.58 deg; joints [-31.343, 12.41, 8.789, -65.592, 42.708, -13.634, -170]
  MoveL 413 to (-2337.75, 783.65, 1090.45) mm, rotated rx -114.42 ry 38.8 rz 164.58 deg; joints [-33.375, 15.887, 5.934, -69.773, 44.392, -10.568, -170]
  MoveL 414 to (-2337.75, 783.65, 1090.45) mm, rotated rx -114.42 ry 38.8 rz 164.58 deg; joints [-33.375, 15.887, 5.934, -69.773, 44.392, -10.568, -170]
  Set speed (50.0 mm/s)
  MoveL 415 to (-2337.75, 790.79, 1070.19) mm, rotated rx -110.09 ry 20.24 rz 173.25 deg; joints [-35.457, 14.134, 5.055, -44.063, 6.364, -24.687, -170]
  MoveL 416 to (-2337.75, 800.76, 1041.89) mm, rotated rx -115.1 ry 36.45 rz 164.18 deg; joints [-33.03, 15.858, 7.052, -67.259, 41.861, -12.102, -170]
  MoveL 417 to (-2337.75, 813.29, 1008.29) mm, rotated rx -105.64 ry 18.04 rz 174.71 deg; joints [-34.546, 14.809, 8.007, -62.538, 19.958, -20.468, -170]
  MoveL 418 to (-2337.75, 823.77, 980.18) mm, rotated rx -101.11 ry 17.55 rz 176.22 deg; joints [-34.184, 15.628, 9.866, -74.944, 30.508, -19.515, -170]
  MoveL 419 to (-2337.75, 836.64, 946.71) mm, rotated rx -101.13 ry 16.53 rz 176.22 deg; joints [-33.895, 15.801, 10.774, -74.768, 30.555, -20.477, -170]
  MoveL 420 to (-2337.75, 847.41, 918.71) mm, rotated rx -101.15 ry 15.69 rz 176.21 deg; joints [-33.648, 15.969, 11.512, -74.606, 30.607, -21.287, -170]
  MoveL 421 to (-2337.75, 847.44, 895.17) mm, rotated rx -98.85 ry 16.34 rz 176.99 deg; joints [-33.639, 16.974, 12.39, -82.131, 37.922, -20.619, -170]
  MoveL 422 to (-2337.75, 847.48, 865.17) mm, rotated rx -95.9 ry 17.72 rz 177.99 deg; joints [-33.666, 18.468, 13.355, -90.749, 47.375, -20.704, -170]
  MoveL 423 to (-2337.75, 847.52, 835.17) mm, rotated rx -92.76 ry 1.83 rz 180 deg; joints [-34.311, 17.71, 12.827, -73.726, 21.892, -33.106, -170]
  MoveL 424 to (-2337.75, 847.55, 805.17) mm, rotated rx -89.9 ry 0.38 rz -179.62 deg; joints [-34.362, 18.852, 13.564, -79.169, 26.454, -34.419, -170]
  MoveL 425 to (-2337.75, 847.49, 781.64) mm, rotated rx -89.88 ry 0.39 rz -179.61 deg; joints [-34.352, 19.451, 13.857, -80.986, 28.333, -34.06, -170]
  MoveL 426 to (-2337.75, 847.4, 751.64) mm, rotated rx -89.85 ry 0.4 rz -179.6 deg; joints [-34.343, 20.233, 14.203, -83.125, 30.619, -33.716, -170]
  MoveL 427 to (-2337.75, 847.31, 721.64) mm, rotated rx -89.82 ry 0.42 rz -179.59 deg; joints [-34.336, 21.038, 14.519, -85.104, 32.806, -33.477, -170]
  MoveL 428 to (-2337.75, 847.23, 691.64) mm, rotated rx -89.79 ry 0.43 rz -179.57 deg; joints [-34.33, 21.864, 14.804, -86.953, 34.912, -33.322, -170]
  MoveL 429 to (-2337.75, 847.13, 668.1) mm, rotated rx -89.79 ry 0.44 rz -179.56 deg; joints [-34.327, 22.523, 15.004, -88.293, 36.481, -33.248, -170]
  MoveL 430 to (-2337.75, 847.01, 638.1) mm, rotated rx -89.78 ry 0.45 rz -179.55 deg; joints [-34.324, 23.382, 15.234, -89.92, 38.429, -33.206, -170]
  MoveL 431 to (-2337.75, 846.89, 608.1) mm, rotated rx -89.77 ry 0.46 rz -179.54 deg; joints [-34.322, 24.26, 15.435, -91.471, 40.326, -33.216, -170]
  MoveL 432 to (-2337.75, 846.77, 578.1) mm, rotated rx -89.76 ry 0.47 rz -179.53 deg; joints [-34.321, 25.158, 15.608, -92.954, 42.178, -33.27, -170]
  MoveL 433 to (-2337.75, 846.63, 534.6) mm, rotated rx -89.77 ry 0.48 rz -179.53 deg; joints [-34.319, 26.487, 15.807, -94.953, 44.742, -33.414, -170]
  MoveL 434 to (-2337.75, 846.54, 504.6) mm, rotated rx -89.78 ry 0.48 rz -179.52 deg; joints [-34.318, 27.425, 15.911, -96.272, 46.468, -33.552, -170]
  MoveL 435 to (-2337.75, 846.44, 474.6) mm, rotated rx -89.79 ry 0.49 rz -179.52 deg; joints [-34.317, 28.381, 15.987, -97.55, 48.16, -33.718, -170]
  MoveL 436 to (-2337.75, 846.34, 444.6) mm, rotated rx -89.79 ry 0.49 rz -179.51 deg; joints [-34.318, 29.354, 16.037, -98.788, 49.822, -33.908, -170]
  MoveL 437 to (-2337.75, 846.24, 414.6) mm, rotated rx -89.8 ry 0.5 rz -179.51 deg; joints [-34.319, 30.344, 16.059, -99.992, 51.454, -34.121, -170]
  MoveL 438 to (-2337.75, 846.15, 384.6) mm, rotated rx -89.81 ry 0.5 rz -179.5 deg; joints [-34.32, 31.349, 16.053, -101.163, 53.058, -34.353, -170]
  MoveL 439 to (-2337.75, 846.05, 354.6) mm, rotated rx -89.81 ry 0.51 rz -179.49 deg; joints [-34.322, 32.37, 16.021, -102.304, 54.634, -34.603, -170]
  MoveL 440 to (-2337.75, 845.95, 324.6) mm, rotated rx -89.82 ry 0.51 rz -179.49 deg; joints [-34.324, 33.405, 15.962, -103.417, 56.183, -34.869, -170]
  MoveL 441 to (-2337.75, 845.85, 294.6) mm, rotated rx -89.83 ry 0.52 rz -179.48 deg; joints [-34.326, 34.454, 15.876, -104.505, 57.706, -35.149, -170]
  MoveL 442 to (-2337.75, 845.76, 264.6) mm, rotated rx -89.83 ry 0.52 rz -179.48 deg; joints [-34.329, 35.517, 15.763, -105.567, 59.202, -35.442, -170]
  MoveL 443 to (-2337.75, 845.66, 234.6) mm, rotated rx -89.84 ry 0.53 rz -179.47 deg; joints [-34.332, 36.593, 15.623, -106.606, 60.673, -35.746, -170]
  MoveL 444 to (-2337.75, 845.56, 204.6) mm, rotated rx -89.85 ry 0.54 rz -179.47 deg; joints [-34.336, 37.681, 15.456, -107.623, 62.118, -36.06, -170]
  MoveL 445 to (-2337.75, 845.54, 196.6) mm, rotated rx -89.85 ry 0.54 rz -179.47 deg; joints [-34.336, 37.973, 15.407, -107.887, 62.497, -36.149, -170]
  Set speed (1000.0 mm/s)
  MoveL 446 to (-2337.75, 845.54, 196.6) mm, rotated rx -89.85 ry 0.54 rz -179.47 deg; joints [-34.336, 37.973, 15.407, -107.887, 62.497, -36.149, -170]
  MoveL 447 to (-2338.67, 945.53, 196.33) mm, rotated rx -89.85 ry 0.54 rz -179.47 deg; joints [-32.082, 35.909, 19.173, -106.286, 64.112, -38.245, -170]
  Set speed (1000.0 mm/s)
  MoveL 448 to (-2418.68, 944.79, 197.17) mm, rotated rx -89.84 ry 0.54 rz -179.46 deg; joints [-34.187, 34.521, 21.849, -110.889, 67.091, -37.41, -170]
  MoveL 449 to (-2417.75, 844.8, 197.45) mm, rotated rx -89.84 ry 0.54 rz -179.46 deg; joints [-36.418, 36.619, 18.026, -112.492, 65.526, -35.305, -170]
  MoveL 450 to (-2417.75, 844.8, 197.45) mm, rotated rx -89.84 ry 0.54 rz -179.46 deg; joints [-36.418, 36.619, 18.026, -112.492, 65.526, -35.305, -170]
  Set speed (50.0 mm/s)
  MoveL 451 to (-2417.75, 844.82, 205.45) mm, rotated rx -89.84 ry 0.54 rz -179.46 deg; joints [-36.417, 36.319, 18.076, -112.236, 65.146, -35.194, -170]
  MoveL 452 to (-2417.75, 844.93, 235.45) mm, rotated rx -89.83 ry 0.53 rz -179.47 deg; joints [-36.41, 35.203, 18.246, -111.242, 63.696, -34.809, -170]
  MoveL 453 to (-2417.75, 845.03, 265.45) mm, rotated rx -89.82 ry 0.53 rz -179.48 deg; joints [-36.405, 34.097, 18.389, -110.242, 62.229, -34.418, -170]
  MoveL 454 to (-2417.75, 845.14, 295.45) mm, rotated rx -89.81 ry 0.52 rz -179.48 deg; joints [-36.4, 33.004, 18.506, -109.224, 60.738, -34.035, -170]
  MoveL 455 to (-2417.75, 845.24, 325.45) mm, rotated rx -89.8 ry 0.51 rz -179.49 deg; joints [-36.396, 31.926, 18.596, -108.188, 59.224, -33.661, -170]
  MoveL 456 to (-2417.75, 845.35, 355.45) mm, rotated rx -89.8 ry 0.51 rz -179.49 deg; joints [-36.392, 30.861, 18.658, -107.132, 57.687, -33.297, -170]
  MoveL 457 to (-2417.75, 845.45, 385.45) mm, rotated rx -89.79 ry 0.5 rz -179.5 deg; joints [-36.389, 29.811, 18.694, -106.056, 56.128, -32.945, -170]
  MoveL 458 to (-2417.75, 845.56, 415.45) mm, rotated rx -89.78 ry 0.5 rz -179.5 deg; joints [-36.385, 28.777, 18.702, -104.957, 54.545, -32.607, -170]
  MoveL 459 to (-2417.75, 845.67, 445.45) mm, rotated rx -89.77 ry 0.49 rz -179.51 deg; joints [-36.383, 27.759, 18.683, -103.836, 52.939, -32.283, -170]
  MoveL 460 to (-2417.75, 845.77, 475.45) mm, rotated rx -89.77 ry 0.49 rz -179.51 deg; joints [-36.38, 26.758, 18.637, -102.689, 51.31, -31.975, -170]
  MoveL 461 to (-2417.75, 845.88, 505.45) mm, rotated rx -89.76 ry 0.48 rz -179.52 deg; joints [-36.378, 25.774, 18.563, -101.516, 49.656, -31.685, -170]
  MoveL 462 to (-2417.75, 845.98, 535.45) mm, rotated rx -89.75 ry 0.48 rz -179.52 deg; joints [-36.377, 24.809, 18.462, -100.313, 47.976, -31.415, -170]
  MoveL 463 to (-2417.75, 846.09, 565.45) mm, rotated rx -89.75 ry 0.47 rz -179.53 deg; joints [-36.376, 23.862, 18.334, -99.078, 46.27, -31.168, -170]
  MoveL 464 to (-2417.75, 846.15, 582.83) mm, rotated rx -89.74 ry 0.47 rz -179.53 deg; joints [-36.375, 23.322, 18.247, -98.346, 45.269, -31.036, -170]
  MoveL 465 to (-2417.75, 846.28, 612.83) mm, rotated rx -89.75 ry 0.46 rz -179.54 deg; joints [-36.373, 22.401, 18.074, -97.018, 43.486, -30.828, -170]
  MoveL 466 to (-2417.75, 846.41, 642.83) mm, rotated rx -89.75 ry 0.45 rz -179.55 deg; joints [-36.372, 21.5, 17.873, -95.645, 41.669, -30.652, -170]
  MoveL 467 to (-2417.75, 846.54, 672.83) mm, rotated rx -89.76 ry 0.44 rz -179.56 deg; joints [-36.371, 20.619, 17.644, -94.221, 39.817, -30.511, -170]
  MoveL 468 to (-2417.75, 846.65, 697.38) mm, rotated rx -89.77 ry 0.43 rz -179.57 deg; joints [-36.371, 19.915, 17.436, -93.012, 38.272, -30.426, -170]
  MoveL 469 to (-2417.75, 846.75, 727.38) mm, rotated rx -89.79 ry 0.42 rz -179.58 deg; joints [-36.372, 19.069, 17.152, -91.433, 36.301, -30.358, -170]
  MoveL 470 to (-2417.75, 846.86, 757.38) mm, rotated rx -89.82 ry 0.41 rz -179.6 deg; joints [-36.373, 18.246, 16.838, -89.773, 34.277, -30.346, -170]
  MoveL 471 to (-2417.75, 846.96, 787.38) mm, rotated rx -89.84 ry 0.39 rz -179.61 deg; joints [-36.376, 17.445, 16.496, -88.015, 32.193, -30.4, -170]
  MoveL 472 to (-2417.75, 847.04, 811.93) mm, rotated rx -89.87 ry 0.38 rz -179.62 deg; joints [-36.38, 16.807, 16.193, -86.49, 30.433, -30.501, -170]
  MoveL 473 to (-2417.75, 847.02, 841.93) mm, rotated rx -92.8 ry 1.7 rz 180 deg; joints [-36.305, 15.603, 15.442, -81.617, 25.936, -28.578, -170]
  MoveL 474 to (-2417.75, 847, 871.93) mm, rotated rx -96.04 ry 17.64 rz 177.94 deg; joints [-35.683, 16.331, 15.914, -94.949, 49.334, -18.274, -170]
  MoveL 475 to (-2417.75, 846.99, 901.93) mm, rotated rx -99.07 ry 16.27 rz 176.91 deg; joints [-35.637, 14.796, 14.931, -86.863, 40.033, -17.596, -170]
  MoveL 476 to (-2417.75, 846.97, 926.49) mm, rotated rx -101.54 ry 15.61 rz 176.08 deg; joints [-35.626, 13.723, 13.997, -79.625, 32.621, -17.705, -170]
  MoveL 477 to (-2417.75, 846.97, 926.49) mm, rotated rx -101.54 ry 15.61 rz 176.08 deg; joints [-35.626, 13.723, 13.997, -79.625, 32.621, -17.705, -170]
  MoveL 478 to (-2417.75, 835.81, 954.33) mm, rotated rx -101.53 ry 16.45 rz 176.08 deg; joints [-35.88, 13.575, 13.232, -79.816, 32.589, -16.845, -170]
  MoveL 479 to (-2417.75, 822.19, 988.31) mm, rotated rx -101.52 ry 17.49 rz 176.09 deg; joints [-36.185, 13.424, 12.274, -80.023, 32.56, -15.805, -170]
  MoveL 480 to (-2417.75, 811.29, 1016.26) mm, rotated rx -106.22 ry 17.96 rz 174.52 deg; joints [-36.525, 12.609, 10.352, -68.881, 22.503, -15.607, -170]
  MoveL 481 to (-2417.75, 798, 1050.37) mm, rotated rx -116.13 ry 36.2 rz 163.55 deg; joints [-35.005, 13.544, 9.297, -68.642, 41.081, -9.503, -170]
  MoveL 482 to (-2417.75, 787.59, 1078.51) mm, rotated rx -115.77 ry 37.52 rz 163.77 deg; joints [-35.22, 13.564, 8.628, -70.021, 42.449, -8.601, -170]
  MoveL 483 to (-2417.75, 779.85, 1099.45) mm, rotated rx -111.03 ry 20.13 rz 172.95 deg; joints [-37.633, 11.908, 6.413, -49.014, 6.917, -19.394, -170]
  MoveL 484 to (-2417.75, 779.74, 1099.76) mm, rotated rx -111.02 ry 20.14 rz 172.95 deg; joints [-37.632, 11.908, 6.411, -49.183, 7.034, -19.296, -170]
  Set speed (1000.0 mm/s)
  MoveL 485 to (-2417.75, 779.74, 1099.76) mm, rotated rx -111.02 ry 20.14 rz 172.95 deg; joints [-37.632, 11.908, 6.411, -49.183, 7.034, -19.296, -170]
  MoveL 486 to (-2418.54, 873.9, 1133.43) mm, rotated rx -115.51 ry 38.56 rz 163.92 deg; joints [-33.383, 10, 10.916, -66.385, 41.362, -11.109, -170]
  Set speed (1000.0 mm/s)
  MoveL 487 to (-2499.41, 869.59, 1143.27) mm, rotated rx -111.27 ry 21.6 rz 172.86 deg; joints [-37.885, 6.215, 11.659, -55.918, 11.743, -14.444, -170]
  MoveL 488 to (-2497.75, 775.46, 1109.54) mm, rotated rx -111.27 ry 21.6 rz 172.86 deg; joints [-39.608, 10.015, 9.031, -69.23, 19.7, -6.621, -170]
  MoveL 489 to (-2497.75, 775.46, 1109.54) mm, rotated rx -111.27 ry 21.6 rz 172.86 deg; joints [-39.608, 10.015, 9.031, -69.23, 19.7, -6.621, -170]
  Set speed (50.0 mm/s)
  MoveL 490 to (-2497.75, 775.82, 1108.56) mm, rotated rx -111.98 ry 20.06 rz 172.64 deg; joints [-39.686, 9.874, 8.43, -60.552, 12.274, -10.709, -170]
  MoveL 491 to (-2497.75, 784.16, 1087.07) mm, rotated rx -112.38 ry 19.01 rz 172.52 deg; joints [-39.574, 9.829, 8.812, -54.987, 8.254, -14.066, -170]
  MoveL 492 to (-2497.75, 795.01, 1059.1) mm, rotated rx -117.19 ry 35.94 rz 162.92 deg; joints [-37.101, 11.312, 11.346, -70.141, 40.219, -6.715, -170]
  MoveL 493 to (-2497.75, 809.17, 1024.35) mm, rotated rx -106.81 ry 17.88 rz 174.33 deg; joints [-38.638, 10.497, 12.524, -75.252, 25.05, -10.735, -170]
  MoveL 494 to (-2497.75, 820.49, 996.57) mm, rotated rx -101.95 ry 17.43 rz 175.94 deg; joints [-38.318, 11.297, 14.508, -85.196, 34.639, -12.027, -170]
  MoveL 495 to (-2497.75, 834.96, 961.95) mm, rotated rx -101.94 ry 16.37 rz 175.94 deg; joints [-37.998, 11.422, 15.526, -84.954, 34.641, -13.15, -170]
  MoveL 496 to (-2497.75, 846.53, 934.27) mm, rotated rx -101.94 ry 15.53 rz 175.94 deg; joints [-37.736, 11.546, 16.319, -84.733, 34.647, -14.059, -170]
  MoveL 497 to (-2497.75, 846.53, 934.27) mm, rotated rx -101.94 ry 15.53 rz 175.94 deg; joints [-37.736, 11.546, 16.319, -84.733, 34.647, -14.059, -170]
  MoveL 498 to (-2497.75, 846.53, 908.7) mm, rotated rx -99.3 ry 16.21 rz 176.83 deg; joints [-37.766, 12.688, 17.31, -91.665, 42.151, -14.538, -170]
  MoveL 499 to (-2497.75, 846.53, 878.7) mm, rotated rx -95.9 ry -2.33 rz -179.99 deg; joints [-38.553, 11.897, 16.054, -67.796, 9.129, -31.381, -170]
  MoveL 500 to (-2497.75, 846.53, 848.7) mm, rotated rx -92.85 ry 1.56 rz 180 deg; joints [-38.449, 13.568, 17.884, -88.991, 29.678, -24.438, -170]
  MoveL 501 to (-2497.75, 846.53, 818.7) mm, rotated rx -89.83 ry 0.38 rz -179.62 deg; joints [-38.544, 14.836, 18.652, -93.403, 34.177, -26.91, -170]
  MoveL 502 to (-2497.75, 846.43, 793.13) mm, rotated rx -89.81 ry 0.4 rz -179.61 deg; joints [-38.544, 15.514, 18.965, -94.699, 35.853, -27.029, -170]
  MoveL 503 to (-2497.75, 846.31, 763.13) mm, rotated rx -89.79 ry 0.41 rz -179.59 deg; joints [-38.546, 16.332, 19.307, -96.159, 37.78, -27.212, -170]
  MoveL 504 to (-2497.75, 846.2, 733.13) mm, rotated rx -89.76 ry 0.42 rz -179.58 deg; joints [-38.548, 17.173, 19.62, -97.562, 39.67, -27.435, -170]
  MoveL 505 to (-2497.75, 846.08, 703.13) mm, rotated rx -89.74 ry 0.44 rz -179.57 deg; joints [-38.552, 18.038, 19.904, -98.918, 41.527, -27.694, -170]
  MoveL 506 to (-2497.75, 845.95, 677.56) mm, rotated rx -89.73 ry 0.44 rz -179.56 deg; joints [-38.554, 18.789, 20.121, -100.012, 43.055, -27.932, -170]
  MoveL 507 to (-2497.75, 845.81, 647.56) mm, rotated rx -89.73 ry 0.45 rz -179.55 deg; joints [-38.558, 19.691, 20.35, -101.262, 44.823, -28.236, -170]
  MoveL 508 to (-2497.75, 845.66, 617.56) mm, rotated rx -89.72 ry 0.46 rz -179.54 deg; joints [-38.562, 20.614, 20.552, -102.481, 46.568, -28.564, -170]
  MoveL 509 to (-2497.75, 845.52, 587.56) mm, rotated rx -89.72 ry 0.47 rz -179.53 deg; joints [-38.566, 21.558, 20.725, -103.672, 48.29, -28.914, -170]
  MoveL 510 to (-2497.75, 845.44, 566.3) mm, rotated rx -89.73 ry 0.47 rz -179.53 deg; joints [-38.568, 22.236, 20.831, -104.48, 49.476, -29.171, -170]
  MoveL 511 to (-2497.75, 845.33, 536.3) mm, rotated rx -89.73 ry 0.48 rz -179.52 deg; joints [-38.571, 23.21, 20.957, -105.6, 51.133, -29.548, -170]
  MoveL 512 to (-2497.75, 845.21, 506.3) mm, rotated rx -89.74 ry 0.48 rz -179.52 deg; joints [-38.574, 24.202, 21.056, -106.701, 52.77, -29.941, -170]
  MoveL 513 to (-2497.75, 845.1, 476.3) mm, rotated rx -89.75 ry 0.49 rz -179.51 deg; joints [-38.578, 25.214, 21.127, -107.783, 54.389, -30.348, -170]
  MoveL 514 to (-2497.75, 844.99, 446.3) mm, rotated rx -89.76 ry 0.5 rz -179.51 deg; joints [-38.582, 26.243, 21.17, -108.847, 55.988, -30.767, -170]
  MoveL 515 to (-2497.75, 844.87, 416.3) mm, rotated rx -89.77 ry 0.5 rz -179.5 deg; joints [-38.587, 27.29, 21.187, -109.895, 57.569, -31.199, -170]
  MoveL 516 to (-2497.75, 844.76, 386.3) mm, rotated rx -89.77 ry 0.51 rz -179.5 deg; joints [-38.592, 28.353, 21.175, -110.928, 59.13, -31.64, -170]
  MoveL 517 to (-2497.75, 844.65, 356.3) mm, rotated rx -89.78 ry 0.51 rz -179.49 deg; joints [-38.597, 29.432, 21.137, -111.946, 60.673, -32.091, -170]
  MoveL 518 to (-2497.75, 844.54, 326.3) mm, rotated rx -89.79 ry 0.52 rz -179.49 deg; joints [-38.603, 30.527, 21.071, -112.949, 62.196, -32.55, -170]
  MoveL 519 to (-2497.75, 844.42, 296.3) mm, rotated rx -89.8 ry 0.52 rz -179.48 deg; joints [-38.609, 31.636, 20.977, -113.94, 63.7, -33.016, -170]
  MoveL 520 to (-2497.75, 844.31, 266.3) mm, rotated rx -89.81 ry 0.53 rz -179.48 deg; joints [-38.615, 32.758, 20.857, -114.917, 65.184, -33.488, -170]
  MoveL 521 to (-2497.75, 844.2, 236.3) mm, rotated rx -89.81 ry 0.53 rz -179.47 deg; joints [-38.621, 33.894, 20.709, -115.881, 66.647, -33.965, -170]
  MoveL 522 to (-2497.75, 844.08, 206.3) mm, rotated rx -89.82 ry 0.54 rz -179.47 deg; joints [-38.628, 35.042, 20.535, -116.832, 68.089, -34.447, -170]
  MoveL 523 to (-2497.75, 844.05, 198.3) mm, rotated rx -89.82 ry 0.54 rz -179.47 deg; joints [-38.629, 35.351, 20.483, -117.08, 68.469, -34.58, -170]
  Set speed (1000.0 mm/s)
  MoveL 524 to (-2497.75, 844.05, 198.3) mm, rotated rx -89.82 ry 0.54 rz -179.47 deg; joints [-38.629, 35.351, 20.483, -117.08, 68.469, -34.58, -170]
  MoveL 525 to (-2498.67, 944.05, 197.99) mm, rotated rx -89.82 ry 0.54 rz -179.47 deg; joints [-36.435, 33.217, 24.368, -115.5, 69.993, -36.691, -170]
  Set speed (1000.0 mm/s)
  MoveL 526 to (-2578.68, 943.31, 198.83) mm, rotated rx -89.82 ry 0.54 rz -179.46 deg; joints [-38.845, 31.989, 26.732, -120.191, 72.849, -36.022, -170]
  MoveL 527 to (-2577.75, 843.31, 199.15) mm, rotated rx -89.82 ry 0.54 rz -179.46 deg; joints [-40.983, 34.162, 22.779, -121.724, 71.359, -33.908, -170]
  MoveL 528 to (-2577.75, 843.31, 199.15) mm, rotated rx -89.82 ry 0.54 rz -179.46 deg; joints [-40.983, 34.162, 22.779, -121.724, 71.359, -33.908, -170]
  Set speed (50.0 mm/s)
  MoveL 529 to (-2577.75, 843.34, 207.15) mm, rotated rx -89.82 ry 0.54 rz -179.46 deg; joints [-40.981, 33.846, 22.832, -121.482, 70.98, -33.753, -170]
  MoveL 530 to (-2577.75, 843.46, 237.15) mm, rotated rx -89.8 ry 0.53 rz -179.47 deg; joints [-40.971, 32.669, 23.01, -120.551, 69.54, -33.202, -170]
  MoveL 531 to (-2577.75, 843.58, 267.15) mm, rotated rx -89.79 ry 0.53 rz -179.48 deg; joints [-40.963, 31.503, 23.162, -119.62, 68.085, -32.639, -170]
  MoveL 532 to (-2577.75, 843.7, 297.15) mm, rotated rx -89.78 ry 0.52 rz -179.48 deg; joints [-40.956, 30.351, 23.287, -118.682, 66.611, -32.079, -170]
  MoveL 533 to (-2577.75, 843.83, 327.15) mm, rotated rx -89.78 ry 0.52 rz -179.49 deg; joints [-40.949, 29.212, 23.383, -117.734, 65.12, -31.522, -170]
  MoveL 534 to (-2577.75, 843.95, 357.14) mm, rotated rx -89.77 ry 0.51 rz -179.49 deg; joints [-40.942, 28.087, 23.453, -116.779, 63.612, -30.969, -170]
  MoveL 535 to (-2577.75, 844.07, 387.14) mm, rotated rx -89.76 ry 0.51 rz -179.5 deg; joints [-40.935, 26.979, 23.495, -115.816, 62.089, -30.422, -170]
  MoveL 536 to (-2577.75, 844.19, 417.14) mm, rotated rx -89.75 ry 0.5 rz -179.5 deg; joints [-40.929, 25.886, 23.509, -114.844, 60.549, -29.88, -170]
  MoveL 537 to (-2577.75, 844.31, 447.14) mm, rotated rx -89.74 ry 0.5 rz -179.51 deg; joints [-40.923, 24.811, 23.496, -113.863, 58.996, -29.345, -170]
  MoveL 538 to (-2577.75, 844.43, 477.14) mm, rotated rx -89.73 ry 0.49 rz -179.51 deg; joints [-40.917, 23.753, 23.455, -112.874, 57.427, -28.818, -170]
  MoveL 539 to (-2577.75, 844.55, 507.14) mm, rotated rx -89.72 ry 0.49 rz -179.52 deg; joints [-40.912, 22.714, 23.386, -111.876, 55.845, -28.299, -170]
  MoveL 540 to (-2577.75, 844.67, 537.14) mm, rotated rx -89.71 ry 0.48 rz -179.52 deg; joints [-40.907, 21.695, 23.29, -110.868, 54.249, -27.789, -170]
  MoveL 541 to (-2577.75, 844.79, 567.14) mm, rotated rx -89.71 ry 0.48 rz -179.52 deg; joints [-40.902, 20.695, 23.166, -109.849, 52.64, -27.29, -170]
  MoveL 542 to (-2577.75, 844.89, 592.29) mm, rotated rx -89.7 ry 0.47 rz -179.53 deg; joints [-40.899, 19.873, 23.041, -108.987, 51.28, -26.88, -170]
  MoveL 543 to (-2577.75, 845.05, 622.29) mm, rotated rx -89.7 ry 0.46 rz -179.54 deg; joints [-40.892, 18.906, 22.866, -107.92, 49.618, -26.397, -170]
  MoveL 544 to (-2577.75, 845.2, 652.29) mm, rotated rx -89.71 ry 0.45 rz -179.55 deg; joints [-40.886, 17.961, 22.664, -106.838, 47.941, -25.929, -170]
  MoveL 545 to (-2577.75, 845.36, 682.29) mm, rotated rx -89.71 ry 0.45 rz -179.56 deg; joints [-40.881, 17.038, 22.434, -105.741, 46.25, -25.476, -170]
  MoveL 546 to (-2577.75, 845.5, 708.87) mm, rotated rx -89.71 ry 0.44 rz -179.56 deg; joints [-40.876, 16.24, 22.207, -104.753, 44.739, -25.089, -170]
  MoveL 547 to (-2577.75, 845.63, 738.87) mm, rotated rx -89.73 ry 0.42 rz -179.58 deg; joints [-40.871, 15.357, 21.921, -103.59, 42.983, -24.659, -170]
  MoveL 548 to (-2577.75, 845.77, 768.87) mm, rotated rx -89.76 ry 0.41 rz -179.59 deg; joints [-40.865, 14.498, 21.607, -102.402, 41.209, -24.251, -170]
  MoveL 549 to (-2577.75, 845.9, 798.87) mm, rotated rx -89.78 ry 0.4 rz -179.6 deg; joints [-40.861, 13.663, 21.266, -101.186, 39.416, -23.868, -170]
  MoveL 550 to (-2577.75, 846.02, 825.46) mm, rotated rx -89.8 ry 0.39 rz -179.61 deg; joints [-40.857, 12.945, 20.94, -100.082, 37.808, -23.551, -170]
  MoveL 551 to (-2577.75, 846.04, 855.46) mm, rotated rx -92.91 ry 1.43 rz 180 deg; joints [-40.745, 11.614, 20.154, -96.089, 33.283, -20.552, -170]
  MoveL 552 to (-2577.75, 846.05, 885.46) mm, rotated rx -96.04 ry -2.41 rz -179.99 deg; joints [-40.73, 9.912, 18.499, -82.859, 17.474, -22.402, -170]
  MoveL 553 to (-2577.75, 846.07, 915.46) mm, rotated rx -99.54 ry 16.15 rz 176.75 deg; joints [-40.036, 10.657, 19.526, -96.583, 44.326, -11.431, -170]
  MoveL 554 to (-2577.75, 846.09, 942.04) mm, rotated rx -102.37 ry 15.45 rz 175.8 deg; joints [-39.985, 9.447, 18.475, -89.989, 36.744, -10.328, -170]
  MoveL 555 to (-2577.75, 834.1, 969.55) mm, rotated rx -102.37 ry 16.28 rz 175.8 deg; joints [-40.252, 9.35, 17.652, -90.238, 36.767, -9.375, -170]
  MoveL 556 to (-2577.75, 818.67, 1004.95) mm, rotated rx -102.38 ry 17.37 rz 175.8 deg; joints [-40.589, 9.259, 16.566, -90.517, 36.798, -8.166, -170]
  MoveL 557 to (-2577.75, 806.92, 1032.55) mm, rotated rx -107.4 ry 17.8 rz 174.13 deg; joints [-40.89, 8.481, 14.52, -81.737, 27.678, -5.823, -170]
  MoveL 558 to (-2577.75, 791.78, 1068.08) mm, rotated rx -113.83 ry 17.65 rz 172.06 deg; joints [-41.556, 7.828, 11.242, -61.228, 9.636, -8.641, -170]
  MoveL 559 to (-2577.75, 780.46, 1095.87) mm, rotated rx -113.38 ry 18.87 rz 172.2 deg; joints [-41.756, 7.888, 10.659, -66.464, 13.462, -5.385, -170]
  MoveL 560 to (-2577.75, 771.44, 1118.01) mm, rotated rx -113.04 ry 19.88 rz 172.3 deg; joints [-41.929, 7.951, 10.162, -69.648, 15.953, -3.382, -170]
  MoveL 561 to (-2577.75, 770.76, 1119.8) mm, rotated rx -112.99 ry 19.98 rz 172.32 deg; joints [-41.941, 7.957, 10.132, -69.976, 16.227, -3.203, -170]
  Set speed (1000.0 mm/s)
  MoveL 562 to (-2577.75, 770.76, 1119.8) mm, rotated rx -112.99 ry 19.98 rz 172.32 deg; joints [-41.941, 7.957, 10.132, -69.976, 16.227, -3.203, -170]
  MoveL 563 to (-2578.66, 863.78, 1156.51) mm, rotated rx -117.81 ry 38.1 rz 162.54 deg; joints [-37.88, 5.461, 14.53, -68.42, 38.462, -5.353, -170]
  Set speed (1000.0 mm/s)
  MoveL 564 to (-2659.56, 858.45, 1167.65) mm, rotated rx -113.47 ry 21.31 rz 172.15 deg; joints [-42.709, 2.254, 14.719, -72.739, 17.68, 0.03, -170]
  MoveL 565 to (-2657.75, 765.6, 1130.54) mm, rotated rx -111.81 ry 2.82 rz 179.99 deg; joints [-45.776, 5.996, 9.604, -106.083, 17.077, 19.354, -170]
  MoveL 566 to (-2657.75, 765.6, 1130.54) mm, rotated rx -111.81 ry 2.82 rz 179.99 deg; joints [-45.776, 5.996, 9.604, -106.083, 17.077, 19.354, -170]
  Set speed (50.0 mm/s)
  MoveL 567 to (-2657.75, 766.69, 1127.82) mm, rotated rx -112.53 ry 1.5 rz 180 deg; joints [-45.681, 6.01, 9.19, -105.676, 14.892, 20.163, -170]
  MoveL 568 to (-2657.75, 776.49, 1104.91) mm, rotated rx -113.06 ry 0.38 rz 180 deg; joints [-45.411, 5.935, 9.685, -103.403, 12.547, 18.966, -170]
  MoveL 569 to (-2657.75, 788.29, 1077.32) mm, rotated rx -113.6 ry -0.75 rz -180 deg; joints [-45.09, 5.859, 10.313, -99.703, 9.436, 16.819, -170]
  MoveL 570 to (-2657.75, 804.52, 1040.87) mm, rotated rx -107.12 ry -1.36 rz -180 deg; joints [-44.349, 5.728, 13.437, -86.135, 6.186, -0.829, -170]
  MoveL 571 to (-2657.75, 816.72, 1013.46) mm, rotated rx -102.26 ry -2.22 rz -180 deg; joints [-43.868, 5.943, 15.716, -84.888, 9.125, -8.937, -170]
  MoveL 572 to (-2657.75, 833.24, 977.13) mm, rotated rx -102.32 ry -3.34 rz -179.99 deg; joints [-43.506, 5.928, 16.691, -76.955, 4.226, -14.611, -170]
  MoveL 573 to (-2657.75, 845.65, 949.82) mm, rotated rx -102.8 ry 15.36 rz 175.65 deg; joints [-42.379, 7.436, 20.463, -95.436, 38.965, -6.508, -170]
  MoveL 574 to (-2657.75, 845.62, 922.22) mm, rotated rx -99.42 ry -3.64 rz -179.99 deg; joints [-43.133, 6.82, 19.122, -85.618, 13.52, -15.248, -170]
  MoveL 575 to (-2657.75, 845.58, 892.22) mm, rotated rx -96.19 ry -2.48 rz -179.99 deg; joints [-43.132, 8.019, 20.675, -93.975, 23.49, -15.957, -170]
  MoveL 576 to (-2657.75, 845.54, 862.22) mm, rotated rx -92.96 ry 1.3 rz 180 deg; joints [-43.196, 9.749, 22.248, -103.047, 36.858, -16.858, -170]
  MoveL 577 to (-2657.75, 845.5, 832.22) mm, rotated rx -89.77 ry 0.39 rz -179.61 deg; joints [-43.324, 11.143, 23.054, -106.638, 41.409, -20.373, -170]
  MoveL 578 to (-2657.75, 845.37, 804.62) mm, rotated rx -89.75 ry 0.4 rz -179.6 deg; joints [-43.329, 11.902, 23.393, -107.573, 42.956, -20.874, -170]
  MoveL 579 to (-2657.75, 845.22, 774.62) mm, rotated rx -89.73 ry 0.42 rz -179.59 deg; joints [-43.336, 12.752, 23.736, -108.581, 44.63, -21.433, -170]
  MoveL 580 to (-2657.75, 845.07, 744.62) mm, rotated rx -89.71 ry 0.43 rz -179.57 deg; joints [-43.342, 13.627, 24.052, -109.582, 46.297, -22.004, -170]
  MoveL 581 to (-2657.75, 844.92, 714.62) mm, rotated rx -89.69 ry 0.44 rz -179.56 deg; joints [-43.35, 14.528, 24.34, -110.576, 47.957, -22.588, -170]
  MoveL 582 to (-2657.75, 844.77, 687.02) mm, rotated rx -89.69 ry 0.45 rz -179.55 deg; joints [-43.355, 15.374, 24.577, -111.463, 49.45, -23.123, -170]
  MoveL 583 to (-2657.75, 844.6, 657.02) mm, rotated rx -89.68 ry 0.46 rz -179.54 deg; joints [-43.362, 16.317, 24.809, -112.424, 51.066, -23.713, -170]
  MoveL 584 to (-2657.75, 844.43, 627.02) mm, rotated rx -89.68 ry 0.47 rz -179.54 deg; joints [-43.369, 17.283, 25.013, -113.38, 52.675, -24.313, -170]
  MoveL 585 to (-2657.75, 844.26, 597.02) mm, rotated rx -89.68 ry 0.48 rz -179.53 deg; joints [-43.377, 18.271, 25.189, -114.334, 54.277, -24.921, -170]
  MoveL 586 to (-2657.75, 844.14, 567.99) mm, rotated rx -89.69 ry 0.48 rz -179.52 deg; joints [-43.382, 19.244, 25.334, -115.231, 55.795, -25.511, -170]
  MoveL 587 to (-2657.75, 844.01, 537.99) mm, rotated rx -89.7 ry 0.48 rz -179.52 deg; joints [-43.388, 20.269, 25.456, -116.155, 57.355, -26.126, -170]
  MoveL 588 to (-2657.75, 843.88, 507.99) mm, rotated rx -89.71 ry 0.49 rz -179.51 deg; joints [-43.394, 21.316, 25.55, -117.078, 58.908, -26.748, -170]
  MoveL 589 to (-2657.75, 843.75, 477.99) mm, rotated rx -89.71 ry 0.49 rz -179.51 deg; joints [-43.4, 22.382, 25.616, -117.999, 60.452, -27.374, -170]
  MoveL 590 to (-2657.75, 843.63, 447.99) mm, rotated rx -89.72 ry 0.5 rz -179.5 deg; joints [-43.407, 23.467, 25.655, -118.918, 61.987, -28.006, -170]
  MoveL 591 to (-2657.75, 843.5, 417.99) mm, rotated rx -89.73 ry 0.5 rz -179.5 deg; joints [-43.414, 24.571, 25.666, -119.835, 63.511, -28.642, -170]
  MoveL 592 to (-2657.75, 843.37, 387.99) mm, rotated rx -89.74 ry 0.51 rz -179.49 deg; joints [-43.422, 25.692, 25.648, -120.749, 65.024, -29.281, -170]
  MoveL 593 to (-2657.75, 843.24, 357.99) mm, rotated rx -89.75 ry 0.51 rz -179.49 deg; joints [-43.43, 26.83, 25.603, -121.661, 66.524, -29.924, -170]
  MoveL 594 to (-2657.75, 843.11, 327.99) mm, rotated rx -89.76 ry 0.52 rz -179.48 deg; joints [-43.438, 27.984, 25.53, -122.57, 68.012, -30.568, -170]
  MoveL 595 to (-2657.75, 842.99, 297.99) mm, rotated rx -89.77 ry 0.52 rz -179.48 deg; joints [-43.446, 29.152, 25.429, -123.475, 69.487, -31.215, -170]
  MoveL 596 to (-2657.75, 842.86, 267.99) mm, rotated rx -89.78 ry 0.53 rz -179.47 deg; joints [-43.455, 30.335, 25.301, -124.377, 70.946, -31.863, -170]
  MoveL 597 to (-2657.75, 842.73, 237.99) mm, rotated rx -89.79 ry 0.53 rz -179.47 deg; joints [-43.464, 31.531, 25.145, -125.275, 72.39, -32.511, -170]
  MoveL 598 to (-2657.75, 842.6, 208) mm, rotated rx -89.8 ry 0.54 rz -179.47 deg; joints [-43.473, 32.74, 24.961, -126.168, 73.817, -33.159, -170]
  MoveL 599 to (-2657.75, 842.57, 200) mm, rotated rx -89.8 ry 0.54 rz -179.47 deg; joints [-43.475, 33.064, 24.907, -126.403, 74.194, -33.336, -170]
  Set speed (1000.0 mm/s)
  MoveL 600 to (-2657.75, 842.57, 200) mm, rotated rx -89.8 ry 0.54 rz -179.47 deg; joints [-43.475, 33.064, 24.907, -126.403, 74.194, -33.336, -170]
  MoveL 601 to (-2658.68, 942.56, 199.65) mm, rotated rx -89.8 ry 0.54 rz -179.47 deg; joints [-41.412, 30.851, 28.929, -124.945, 75.657, -35.452, -170]
  Set speed (1000.0 mm/s)
  MoveL 602 to (-2738.68, 941.82, 200.49) mm, rotated rx -89.79 ry -19.46 rz -179.53 deg; joints [-43.229, 25.653, 30.46, -100.805, 39.565, -43.756, -170]
  MoveL 603 to (-2737.75, 841.82, 200.86) mm, rotated rx -89.8 ry 0.54 rz -179.46 deg; joints [-46.117, 32.05, 26.864, -131.171, 76.992, -32.797, -170]
  MoveL 604 to (-2737.75, 841.82, 200.86) mm, rotated rx -89.8 ry 0.54 rz -179.46 deg; joints [-46.117, 32.05, 26.864, -131.171, 76.992, -32.797, -170]
  Set speed (50.0 mm/s)
  MoveL 605 to (-2737.75, 841.85, 208.85) mm, rotated rx -89.8 ry 0.54 rz -179.46 deg; joints [-46.114, 31.718, 26.919, -130.943, 76.619, -32.599, -170]
  MoveL 606 to (-2737.75, 841.99, 238.85) mm, rotated rx -89.78 ry 0.53 rz -179.47 deg; joints [-46.102, 30.483, 27.107, -130.072, 75.206, -31.885, -170]
  MoveL 607 to (-2737.75, 842.13, 268.84) mm, rotated rx -89.77 ry 0.53 rz -179.47 deg; joints [-46.092, 29.258, 27.268, -129.207, 73.781, -31.152, -170]
  MoveL 608 to (-2737.75, 842.27, 298.84) mm, rotated rx -89.76 ry 0.52 rz -179.48 deg; joints [-46.082, 28.046, 27.4, -128.342, 72.341, -30.418, -170]
  MoveL 609 to (-2737.75, 842.4, 328.84) mm, rotated rx -89.75 ry 0.52 rz -179.48 deg; joints [-46.073, 26.848, 27.505, -127.477, 70.89, -29.683, -170]
  MoveL 610 to (-2737.75, 842.54, 358.84) mm, rotated rx -89.74 ry 0.51 rz -179.49 deg; joints [-46.064, 25.665, 27.582, -126.614, 69.427, -28.948, -170]
  MoveL 611 to (-2737.75, 842.67, 388.84) mm, rotated rx -89.73 ry 0.51 rz -179.49 deg; joints [-46.055, 24.499, 27.63, -125.752, 67.955, -28.212, -170]
  MoveL 612 to (-2737.75, 842.81, 418.84) mm, rotated rx -89.72 ry 0.51 rz -179.5 deg; joints [-46.047, 23.35, 27.65, -124.893, 66.473, -27.478, -170]
  MoveL 613 to (-2737.75, 842.94, 448.84) mm, rotated rx -89.71 ry 0.5 rz -179.5 deg; joints [-46.039, 22.219, 27.642, -124.037, 64.984, -26.744, -170]
  MoveL 614 to (-2737.75, 843.08, 478.84) mm, rotated rx -89.7 ry 0.5 rz -179.51 deg; joints [-46.032, 21.106, 27.606, -123.185, 63.488, -26.011, -170]
  MoveL 615 to (-2737.75, 843.21, 508.84) mm, rotated rx -89.69 ry 0.49 rz -179.51 deg; joints [-46.024, 20.013, 27.542, -122.337, 61.986, -25.281, -170]
  MoveL 616 to (-2737.75, 843.35, 538.84) mm, rotated rx -89.68 ry 0.49 rz -179.52 deg; joints [-46.018, 18.941, 27.449, -121.494, 60.48, -24.552, -170]
  MoveL 617 to (-2737.75, 843.48, 568.84) mm, rotated rx -89.67 ry 0.48 rz -179.52 deg; joints [-46.011, 17.89, 27.329, -120.656, 58.971, -23.826, -170]
  MoveL 618 to (-2737.75, 843.63, 601.75) mm, rotated rx -89.66 ry 0.48 rz -179.53 deg; joints [-46.004, 16.763, 27.165, -119.744, 57.312, -23.033, -170]
  MoveL 619 to (-2737.75, 843.81, 631.75) mm, rotated rx -89.66 ry 0.47 rz -179.53 deg; joints [-45.996, 15.753, 26.986, -118.896, 55.773, -22.307, -170]
  MoveL 620 to (-2737.75, 843.99, 661.75) mm, rotated rx -89.66 ry 0.46 rz -179.54 deg; joints [-45.988, 14.767, 26.78, -118.054, 54.233, -21.584, -170]
  MoveL 621 to (-2737.75, 844.17, 691.75) mm, rotated rx -89.66 ry 0.45 rz -179.55 deg; joints [-45.981, 13.806, 26.547, -117.219, 52.692, -20.866, -170]
  MoveL 622 to (-2737.75, 844.35, 720.36) mm, rotated rx -89.66 ry 0.44 rz -179.56 deg; joints [-45.974, 12.911, 26.298, -116.429, 51.224, -20.184, -170]
  MoveL 623 to (-2737.75, 844.51, 750.36) mm, rotated rx -89.68 ry 0.43 rz -179.57 deg; joints [-45.966, 11.995, 26.007, -115.585, 49.657, -19.461, -170]
  MoveL 624 to (-2737.75, 844.67, 780.36) mm, rotated rx -89.7 ry 0.42 rz -179.58 deg; joints [-45.959, 11.104, 25.689, -114.748, 48.091, -18.743, -170]
  MoveL 625 to (-2737.75, 844.83, 810.36) mm, rotated rx -89.72 ry 0.41 rz -179.6 deg; joints [-45.952, 10.24, 25.344, -113.919, 46.529, -18.03, -170]
  MoveL 626 to (-2737.75, 844.99, 838.98) mm, rotated rx -89.73 ry 0.39 rz -179.61 deg; joints [-45.946, 9.441, 24.989, -113.135, 45.042, -17.355, -170]
  MoveL 627 to (-2737.75, 845.05, 868.98) mm, rotated rx -93.02 ry 1.16 rz 180 deg; joints [-45.805, 7.984, 24.163, -109.94, 40.475, -13.331, -170]
  MoveL 628 to (-2737.75, 845.1, 898.98) mm, rotated rx -96.34 ry -2.55 rz -179.99 deg; joints [-45.719, 6.229, 22.634, -103.684, 28.787, -10.535, -170]
  MoveL 629 to (-2737.75, 845.16, 928.98) mm, rotated rx -99.66 ry -3.69 rz -179.99 deg; joints [-45.688, 5.017, 21.163, -99.681, 21.453, -7.029, -170]
  MoveL 630 to (-2737.75, 845.21, 957.6) mm, rotated rx -102.81 ry -4.22 rz -179.99 deg; joints [-45.701, 4.109, 19.68, -96.687, 15.623, -3.405, -170]
  MoveL 631 to (-2737.75, 832.36, 984.71) mm, rotated rx -102.76 ry -3.39 rz -179.99 deg; joints [-46.02, 4.134, 18.837, -99.386, 17.301, -1.104, -170]
  MoveL 632 to (-2737.75, 814.63, 1022.1) mm, rotated rx -102.71 ry -2.25 rz -179.99 deg; joints [-46.452, 4.204, 17.634, -102.624, 19.358, 1.78, -170]
  MoveL 633 to (-2737.75, 801.97, 1049.3) mm, rotated rx -107.7 ry -1.38 rz -180 deg; joints [-46.969, 4.062, 15.342, -107.23, 18.678, 11.904, -170]
  MoveL 634 to (-2737.75, 784.5, 1086.82) mm, rotated rx -114.59 ry -0.74 rz -180 deg; joints [-47.844, 4.334, 11.839, -118.897, 20.974, 28.637, -170]
  MoveL 635 to (-2737.75, 772.22, 1114.19) mm, rotated rx -114.09 ry 0.37 rz 180 deg; joints [-48.171, 4.452, 11.089, -120.27, 22.649, 29.451, -170]
  MoveL 636 to (-2737.75, 761.54, 1137.99) mm, rotated rx -113.67 ry 1.37 rz 180 deg; joints [-48.448, 4.569, 10.425, -121.258, 24.016, 30.053, -170]
  MoveL 637 to (-2737.75, 759.94, 1141.75) mm, rotated rx -113.56 ry 1.56 rz 180 deg; joints [-48.49, 4.584, 10.339, -121.34, 24.24, 30.061, -170]
  Set speed (1000.0 mm/s)
  MoveL 638 to (-2737.75, 759.94, 1141.75) mm, rotated rx -113.56 ry 1.56 rz 180 deg; joints [-48.49, 4.584, 10.339, -121.34, 24.24, 30.061, -170]
  MoveL 639 to (-2738.83, 851.61, 1181.71) mm, rotated rx -113.56 ry 1.56 rz 180 deg; joints [-46.899, 0.555, 12.87, -115.16, 18.964, 28.183, -170]
  Set speed (1000.0 mm/s)
  MoveL 640 to (-2819.7, 845.03, 1194.22) mm, rotated rx -114.09 ry 2.76 rz 179.99 deg; joints [-50.084, -0.832, 14.225, -128.62, 28.917, 35.737, -170]
  MoveL 641 to (-2817.75, 753.74, 1153.45) mm, rotated rx -114.09 ry 2.76 rz 179.99 deg; joints [-51.484, 3.298, 11.616, -132.022, 32.557, 35.842, -170]
  MoveL 642 to (-2817.75, 753.74, 1153.45) mm, rotated rx -114.09 ry 2.76 rz 179.99 deg; joints [-51.484, 3.298, 11.616, -132.022, 32.557, 35.842, -170]
  Set speed (50.0 mm/s)
  MoveL 643 to (-2817.75, 755.95, 1148.51) mm, rotated rx -114.64 ry 1.63 rz 180 deg; joints [-51.376, 3.296, 11.426, -132.884, 31.643, 36.99, -170]
  MoveL 644 to (-2817.75, 767.63, 1123.72) mm, rotated rx -115.16 ry 0.36 rz 180 deg; joints [-51.07, 3.14, 12.1, -132.55, 30.318, 36.883, -170]
  MoveL 645 to (-2817.75, 780.41, 1096.58) mm, rotated rx -115.61 ry -0.73 rz -180 deg; joints [-50.743, 2.977, 12.924, -131.75, 29, 36.347, -170]
  MoveL 646 to (-2817.75, 799.26, 1057.85) mm, rotated rx -108.27 ry -1.39 rz -180 deg; joints [-49.789, 2.539, 16.794, -120.245, 26.501, 19.504, -170]
